// TwinCAT 3 PLC project PLC_Tank
// ProgramVersion: 3.1.4026.27
// libraries:
//   Tc2_ControllerToolbox, * (Beckhoff Automation GmbH)
//   Tc2_ModbusSrv, * (Beckhoff Automation GmbH)
//   Tc2_Standard, * (Beckhoff Automation GmbH)
//   Tc2_System, * (Beckhoff Automation GmbH)
//   Tc3_Module, * (Beckhoff Automation GmbH)
//   VisuDialogs, * (System)
//   VisuSymbols,newest,System
// project tree:
//   DUTs/ TAnalogConversion.TcDUT, TEngine.TcDUT, TEngineCmd.TcDUT, THeaterState.TcDUT, THeaterCmd.TcDUT, THeater.TcDUT, TPhaseHeating.TcDUT, TPhaseCmd.TcDUT, TPhaseDraining.TcDUT, TPhaseFilling.TcDUT, TPhaseMixing.TcDUT, TPhaseState.TcDUT, TValveState.TcDUT, TValveCmd.TcDUT, TEngineState.TcDUT, TTank.TcDUT, TValve.TcDUT
//   / GlobalTextList.TcGTLO, PlcTask.TcTTO, PlcTask500ms.TcTTO, Visualization Manager.TcVMO (not stored)
//   GVLs/ Global.TcGVL
//   POUs/ Draining.TcPOU, Engine_1DO.TcPOU, FB_Tank.TcPOU, Filling.TcPOU, Heater.TcPOU, Heating.TcPOU, Main_Batch.TcPOU, MB_Connector.TcPOU, Mixing.TcPOU, Test.TcPOU, Valve_2DO.TcPOU, MAIN.TcPOU
//   POUs/Misc/ EngToRaw.TcPOU, RawToEng.TcPOU
//   VISUs/ Visualization.TcVIS
// real-time tasks:
//   TASK PlcTask: cycle T#100000us, priority 20, ADS port 350
//   TASK PlcTask500ms: cycle T#500ms, priority 1, ADS port 351

CONFIGURATION PLC_Tank
    RESOURCE PLC ON TwinCAT3
        TASK PlcTask(INTERVAL := T#100000us, PRIORITY := 20);
        TASK PlcTask500ms(INTERVAL := T#500ms, PRIORITY := 1);
        PROGRAM MB_Connector WITH PlcTask : MB_Connector;
        PROGRAM Main_Batch WITH PlcTask : Main_Batch;
        PROGRAM MAIN WITH PlcTask500ms : MAIN;
    END_RESOURCE
END_CONFIGURATION

// ---- DUTs/TAnalogConversion.TcDUT
TYPE TAnalogConversion :
STRUCT
	TransducerLoLevel : UINT;
	TransducerHiLevel : UINT;
	ScaledValLoLevel : REAL;
	ScaledValHiLevel : REAL;
END_STRUCT
END_TYPE

// ---- DUTs/TEngine.TcDUT
TYPE TEngine :
STRUCT
	Cmd : TEngineCmd;
	State : TEngineState;
	Time2Start : TIME := T#5S;
	RisingEdgeTrigger : R_TRIG;
	StartupFailTimer : TON;
END_STRUCT
END_TYPE

// ---- DUTs/TEngineCmd.TcDUT
TYPE TEngineCmd :
STRUCT
		SetRT : DINT;
		AutCtrl : BOOL;
		ManCtrl : BOOL;
		TurnOnMan : BOOL;
		TurnOffMan : BOOL;
		Req2RunAutCtrl : BOOL;
		ResetSUF : BOOL;
END_STRUCT
END_TYPE

// ---- DUTs/THeaterState.TcDUT
TYPE THeaterState :
STRUCT
	EnableOut : BOOL;
	HeatingOut : REAL;
	AutCtrl : BOOL;
	ManCtrl : BOOL;
	MayRun : BOOL;
	MayAutoRun : BOOL;
	Err 	: BOOL;
	StateInt : INT;
	GenErr : BOOL; //signalisation: error occured

	HeatingPower : REAL;
	

END_STRUCT
END_TYPE

// ---- DUTs/THeaterCmd.TcDUT
TYPE THeaterCmd :
STRUCT
	AutCtrl : BOOL;
	ManCtrl : BOOL;
	TurnOnMan : BOOL;
	TurnOffMan : BOOL;
	Req2RunAutCtrl : BOOL;
END_STRUCT
END_TYPE

// ---- DUTs/THeater.TcDUT
TYPE THeater :
STRUCT
	Cmd : THeaterCmd;
	State : THeaterState;
	
	ParamHeatingPowerManual : REAL := 50.0;
	ParamHeatingSetPointAutomat : REAL := 60.0;
	
	PID : FB_CTRL_PID;
	ThresholdTimer : TON;
	
END_STRUCT
END_TYPE

// ---- DUTs/TPhaseHeating.TcDUT
TYPE TPhaseHeating :
STRUCT
	Cmd : TPhaseCmd;
	State : TPhaseState;
	
	ParamReqTemp : REAL;
	
	WaterTemp : REAL;
	
	fTime : INT;
END_STRUCT
END_TYPE

// ---- DUTs/TPhaseCmd.TcDUT
TYPE TPhaseCmd :
STRUCT
	StartAut : BOOL;
	StopAut : BOOL;
	StartMan : BOOL;
	StopMan : BOOL;
	PauseMan : BOOL;
	ResumeMan : BOOL;
	ResetDone : BOOL;
	AutCtrl : BOOL;
	ManCtrl : BOOL;
END_STRUCT
END_TYPE

// ---- DUTs/TPhaseDraining.TcDUT
TYPE TPhaseDraining :
STRUCT
	Cmd : TPhaseCmd;
	State : TPhaseState;
	
	ParamDrainLevel : REAL;
	WaterLevel : REAL;
END_STRUCT
END_TYPE

// ---- DUTs/TPhaseFilling.TcDUT
TYPE TPhaseFilling :
STRUCT
	Cmd : TPhaseCmd;
	State : TPhaseState;
	
	ParamFillLevel : REAL;
	WaterLevel : REAL;
END_STRUCT
END_TYPE

// ---- DUTs/TPhaseMixing.TcDUT
TYPE TPhaseMixing :
STRUCT
	Cmd : TPhaseCmd;
	State : TPhaseState;
	
	ParamTimeSec : INT;
	
	ElapsedTimeSec : INT;
END_STRUCT
END_TYPE

// ---- DUTs/TPhaseState.TcDUT
TYPE TPhaseState :
STRUCT
	Running : BOOL;
	Idle : BOOL;
	Paused : BOOL;
	Done : BOOL;
	AutCtrl : BOOL;
	ManCtrl : BOOL;
	Stateint : INT;
END_STRUCT
END_TYPE

// ---- DUTs/TValveState.TcDUT
TYPE TValveState :
STRUCT
		Open : BOOL;
		Closed : BOOL;
		OpenOut : BOOL;
		CloseOut : BOOL;
		Err : BOOL;
		StartupFail : BOOL;
		AutCtrl : BOOL;
		ManCtrl : BOOL;
		MayRun : BOOL;
		MayAutoRun : BOOL; //device is working in automatic regime
		GenErr : BOOL; //signalisation: error occured
		StColor : INT; //valve state: Open(0), Closed(1), OpenAndErr(2), ClosedAndErr(3) ,NotOpenNotClosedNotErr(4), NotOpenNotClosedAndErr(5), OpenAndClosedAndErr(6), OpenAndClosedNotErr(7)

END_STRUCT
END_TYPE

// ---- DUTs/TValveCmd.TcDUT
TYPE TValveCmd :
STRUCT
		AutCtrl : BOOL;
		ManCtrl : BOOL;
		OpenMan : BOOL;
		StopMan : BOOL;
		CloseMan : BOOL;
		Req2OpenAut : BOOL;
		Req2CloseAut : BOOL;
		ResetSUF : BOOL;
END_STRUCT
END_TYPE

// ---- DUTs/TEngineState.TcDUT
TYPE TEngineState :
STRUCT
		RT : DINT;
		Run : BOOL;
		RunOut : BOOL;
		Err : BOOL;
		StartUpFail : BOOL;
		AutCtrl : BOOL;
		ManCtrl : BOOL;
		MayRun : BOOL;
		MayAutoRun : BOOL;
		GenErr : BOOL;
		StateInt : INT;
		
		StartupFailTime : INT;
END_STRUCT
END_TYPE

// ---- DUTs/TTank.TcDUT
TYPE TTank :
STRUCT
	Mixer : TEngine;
	ValveFilling : TValve;
	ValveDraining : TValve;
	Heater : THeater;
	
	Filling : TPhaseFilling;
	Draining : TPhaseDraining;
	Mixing : TPhaseMixing;
	Heating : TPhaseHeating;
	
	GlobalError : BOOL;

END_STRUCT
END_TYPE

// ---- DUTs/TValve.TcDUT
TYPE TValve :
STRUCT
	Cmd : TValveCmd;
	State : TValveState;
	Time2Open : TIME := T#12S;
	
	OpenFailTimer : TON;
	CloseFailTimer : TON;
	
END_STRUCT
END_TYPE

// ---- GVLs/Global.TcGVL
{attribute 'qualified_only'}
VAR_GLOBAL
	Tank1 : TTank;
	

	secImp : BOOL;
	
	diMixerRun : BOOL;
	diMixerError : BOOL;
	diValveFillOpen : BOOL;
	diValveFillClose : BOOL;
	diValveFillError : BOOL;
	diValveDrainOpen : BOOL;
	diValveDrainClose : BOOL;
	diValveDrainError : BOOL;
	
	aiWaterLevel : WORD;
	aiWaterTemp : WORD;
	
	doMixerStart : BOOL;
	doValveFillOpen : BOOL;
	doValveFillClose : BOOL;
	doValveDrainOpen : BOOL;
	doValveDrainClose : BOOL;
	doHeatingEnable : BOOL;
	
	aoReqPowerOfHeating : WORD;

END_VAR

VAR_GLOBAL CONSTANT
	Running : INT := 0;
	Stop : INT := 1;
	RunningAndError : INT := 2;
	Err : INT := 3;

	PhIdle : INT := 0;
	PhRunning : INT := 1;
	PhPause : INT := 2;
	
    Open : INT := 0;
	Closed : INT := 1;
	OpenAndErr : INT := 2;
	ClosedAndErr : INT := 3;
	NotOpenNotClosedNotErr : INT := 4;
	NotOpenNotClosedAndErr : INT := 5;
	OpenAndClosedAndErr : INT := 6;
	OpenAndClosedNotErr : INT := 7;
END_VAR

// ---- POUs/MB_Connector.TcPOU
PROGRAM MB_Connector
VAR
	
    mb_ipaddr   : STRING(15) := '127.0.0.1';
    mb_port     : UINT := 504;
    mb_unitid   : BYTE := 1;
	
	fbReadRegs		: FB_MBReadInputRegs;
	mb_regs    		: ARRAY [0..4] OF WORD;
	mb_regs_error	: BOOL;
	mb_regs_busy	: BOOL;
	mb_regs_execute : BOOL;
	mb_regs_errid	: UDINT;
	
	fbReadInps	: FB_MBReadInputs;
	mb_inps			: ARRAY [0..4] OF BYTE;
	mb_inps_error	: BOOL;
	mb_inps_busy	: BOOL;
	mb_inps_execute : BOOL;
	mb_inps_errid	: UDINT;
	
	fbWriteRegs		: FB_MBWriteRegs;
	mbw_regs    	: ARRAY [0..4] OF WORD;
	mbw_regs_error	: BOOL;
	mbw_regs_busy	: BOOL;
	mbw_regs_execute: BOOL;
	mbw_regs_errid	: UDINT;
	
	fbWriteCoils	: FB_MBWriteCoils;
	mbw_coils		: ARRAY [0..4] OF BYTE;
	mbw_coils_error	: BOOL;
	mbw_coils_busy	: BOOL;
	mbw_coils_execute: BOOL;
	mbw_coils_errid	: UDINT;
	
END_VAR

fbReadRegs.sIPAddr := mb_ipaddr;
fbReadRegs.nTCPPort := mb_port;
fbReadRegs.nQuantity := 4;
fbReadRegs.nMBAddr := 0;
fbReadRegs.cbLength := SIZEOF(mb_regs);
fbReadRegs.pDestAddr := ADR(mb_regs);
fbReadRegs.nUnitID := mb_unitid;
fbReadRegs.tTimeout := T#5S;
IF (mb_regs_busy = FALSE) THEN
	mb_regs_execute := TRUE;
ELSE
	mb_regs_execute := FALSE;
END_IF
fbReadRegs(bExecute := mb_regs_execute, 
		   bBusy => mb_regs_busy, bError => mb_regs_error, 
		   nErrId => mb_regs_errid);



fbReadInps.sIPAddr := mb_ipaddr;
fbReadInps.nTCPPort := mb_port;
fbReadInps.nQuantity := 32;
fbReadInps.nMBAddr := 0;
fbReadInps.cbLength := SIZEOF(mb_inps);
fbReadInps.pDestAddr := ADR(mb_inps);
fbReadInps.nUnitID := mb_unitid;
fbReadInps.tTimeout := T#5S;
IF (mb_inps_busy = FALSE) THEN
	mb_inps_execute := TRUE;
ELSE
	mb_inps_execute := FALSE;
END_IF
fbReadInps(bExecute := mb_inps_execute, 
	bBusy => mb_inps_busy, bError => mb_inps_error, nErrId => mb_inps_errid);

Global.diValveFillOpen := mb_inps[0].0;
Global.diValveFillClose := mb_inps[0].1;
Global.diValveFillError := mb_inps[0].2;
Global.diValveDrainOpen := mb_inps[0].3;
Global.diValveDrainClose := mb_inps[0].4;
Global.diValveDrainError := mb_inps[0].5;
Global.diMixerRun := mb_inps[0].6;
Global.diMixerError := mb_inps[0].7;

Global.aiWaterLevel := mb_regs[0];
Global.aiWaterTemp := mb_regs[2];







fbWriteRegs.sIPAddr := mb_ipaddr;
fbWriteRegs.nTCPPort := mb_port;
fbWriteRegs.nQuantity := 4;
fbWriteRegs.nMBAddr := 0;
fbWriteRegs.cbLength := SIZEOF(mbw_regs);
fbWriteRegs.pSrcAddr := ADR(mbw_regs);
fbWriteRegs.nUnitID := mb_unitid;
fbWriteRegs.tTimeout := T#5S;
IF (mbw_regs_busy = FALSE) THEN
	mbw_regs_execute := TRUE;
ELSE
	mbw_regs_execute := FALSE;
END_IF
fbWriteRegs(bExecute := mbw_regs_execute, 
		   bBusy => mbw_regs_busy, bError => mbw_regs_error, 
		   nErrId => mbw_regs_errid);



fbWriteCoils.sIPAddr := mb_ipaddr;
fbWriteCoils.nTCPPort := mb_port;
fbWriteCoils.nQuantity := 32;
fbWriteCoils.nMBAddr := 0;
fbWriteCoils.cbLength := SIZEOF(mbw_coils);
fbWriteCoils.pSrcAddr := ADR(mbw_coils);
fbWriteCoils.nUnitID := mb_unitid;
fbWriteCoils.tTimeout := T#5S;
IF (mbw_coils_busy = FALSE) THEN
	mbw_coils_execute := TRUE;
ELSE
	mbw_coils_execute := FALSE;
END_IF
fbWriteCoils(bExecute := mbw_coils_execute, 
	bBusy => mbw_coils_busy, bError => mbw_coils_error, nErrId => mbw_coils_errid);

mbw_coils[0].0 := Global.doValveFillOpen;
mbw_coils[0].1 := Global.doValveFillClose;
mbw_coils[0].2 := Global.doValveDrainOpen;
mbw_coils[0].3 := Global.doValveDrainClose;
mbw_coils[0].4 := Global.doMixerStart;
mbw_coils[0].5 := Global.doHeatingEnable;

mbw_regs[0] := Global.aoReqPowerOfHeating;

END_PROGRAM

// ---- POUs/Main_Batch.TcPOU
PROGRAM Main_Batch
VAR
	FB_Tank_1 : FB_Tank;
END_VAR

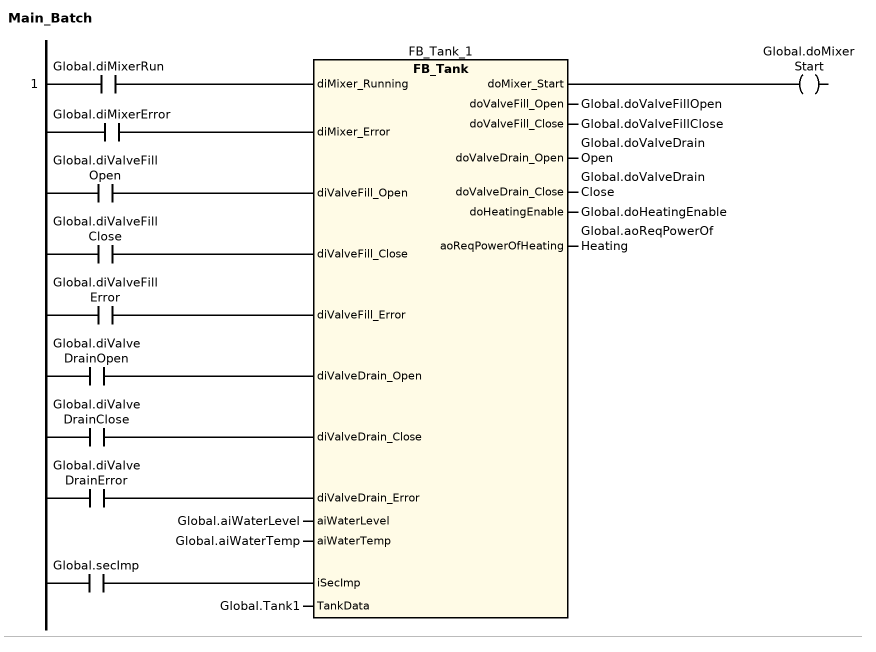
// NETWORK 1
FB_Tank_1(
    diMixer_Running := Global.diMixerRun,
    diMixer_Error := Global.diMixerError,
    diValveFill_Open := Global.diValveFillOpen,
    diValveFill_Close := Global.diValveFillClose,
    diValveFill_Error := Global.diValveFillError,
    diValveDrain_Open := Global.diValveDrainOpen,
    diValveDrain_Close := Global.diValveDrainClose,
    diValveDrain_Error := Global.diValveDrainError,
    aiWaterLevel := Global.aiWaterLevel,
    aiWaterTemp := Global.aiWaterTemp,
    iSecImp := Global.secImp,
    TankData := Global.Tank1,
    doValveFill_Open => Global.doValveFillOpen,
    doValveFill_Close => Global.doValveFillClose,
    doValveDrain_Open => Global.doValveDrainOpen,
    doValveDrain_Close => Global.doValveDrainClose,
    doHeatingEnable => Global.doHeatingEnable,
    aoReqPowerOfHeating => Global.aoReqPowerOfHeating); // FB_Tank
Global.doMixerStart := FB_Tank_1.doMixer_Start;

END_PROGRAM

// ---- POUs/FB_Tank.TcPOU
FUNCTION_BLOCK FB_Tank
VAR_INPUT
	diMixer_Running : BOOL;
	diMixer_Error : BOOL;
	diValveFill_Open : BOOL;
	diValveFill_Close : BOOL;
	diValveFill_Error : BOOL;
	diValveDrain_Open : BOOL;
	diValveDrain_Close : BOOL;
	diValveDrain_Error : BOOL;
	aiWaterLevel : WORD;
	aiWaterTemp : WORD;
	iSecImp : BOOL; //Požaduje se vstup s periodou 1 sekunda a libovolnou střídou
END_VAR

VAR_OUTPUT
	doMixer_Start : BOOL;
	doValveFill_Open : BOOL;
	doValveFill_Close : BOOL;
	doValveDrain_Open : BOOL;
	doValveDrain_Close : BOOL;
	doHeatingEnable : BOOL;
	aoReqPowerOfHeating : WORD;
END_VAR

VAR_IN_OUT
	TankData : TTank;
END_VAR

VAR
	//Konfigurace přepočtu rozsahu převodníků
	WaterTemp : TAnalogConversion := (TransducerLoLevel := 0, TransducerHiLevel := 27648, ScaledValLoLevel := 0, ScaledValHiLevel := 100);
	WaterLevel : TAnalogConversion := (TransducerLoLevel := 0, TransducerHiLevel := 27648, ScaledValLoLevel := 0, ScaledValHiLevel := 2);
	ReqOutputPower : TAnalogConversion := (ScaledValLoLevel := 0, ScaledValHiLevel := 100, TransducerLoLevel := 0, TransducerHiLevel := 27648);

	//Instance zanořených funkčních bloků
	ValveDrainCm : Valve_2DO;
	ValveFillCm : Valve_2DO;
	MixerCm : Engine_1DO;
	HeaterCm : Heater;
	FillingPhase : Filling;
	MixingPhase : Mixing;
	DrainingPhase : Draining;
	HeatingPhase : Heating;
	TON1: TON;
	RawToEng_1: RawToEng;
	RawToEng_2: RawToEng;
	EngToRaw_1: EngToRaw;
END_VAR

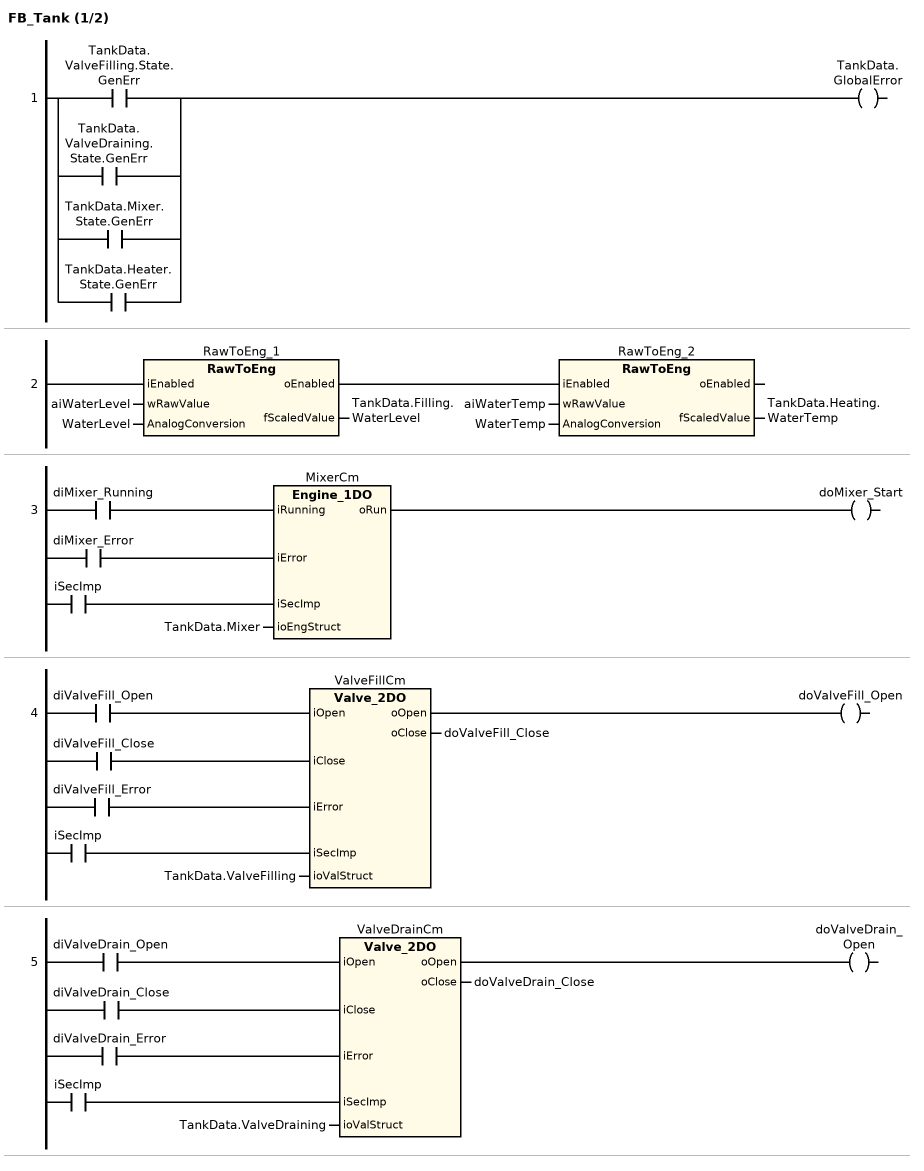
// NETWORK 1
TankData.GlobalError := TankData.ValveFilling.State.GenErr OR TankData.ValveDraining.State.GenErr OR TankData.Mixer.State.GenErr OR TankData.Heater.State.GenErr;

// NETWORK 2
RawToEng_1(
    iEnabled := TRUE,
    wRawValue := aiWaterLevel,
    AnalogConversion := WaterLevel,
    fScaledValue => TankData.Filling.WaterLevel); // RawToEng
RawToEng_2(
    iEnabled := RawToEng_1.oEnabled,
    wRawValue := aiWaterTemp,
    AnalogConversion := WaterTemp,
    fScaledValue => TankData.Heating.WaterTemp); // RawToEng

// NETWORK 3
MixerCm(
    iRunning := diMixer_Running,
    iError := diMixer_Error,
    iSecImp := iSecImp,
    ioEngStruct := TankData.Mixer); // Engine_1DO
doMixer_Start := MixerCm.oRun;

// NETWORK 4
ValveFillCm(
    iOpen := diValveFill_Open,
    iClose := diValveFill_Close,
    iError := diValveFill_Error,
    iSecImp := iSecImp,
    ioValStruct := TankData.ValveFilling,
    oClose => doValveFill_Close); // Valve_2DO
doValveFill_Open := ValveFillCm.oOpen;

// NETWORK 5
ValveDrainCm(
    iOpen := diValveDrain_Open,
    iClose := diValveDrain_Close,
    iError := diValveDrain_Error,
    iSecImp := iSecImp,
    ioValStruct := TankData.ValveDraining,
    oClose => doValveDrain_Close); // Valve_2DO
doValveDrain_Open := ValveDrainCm.oOpen;

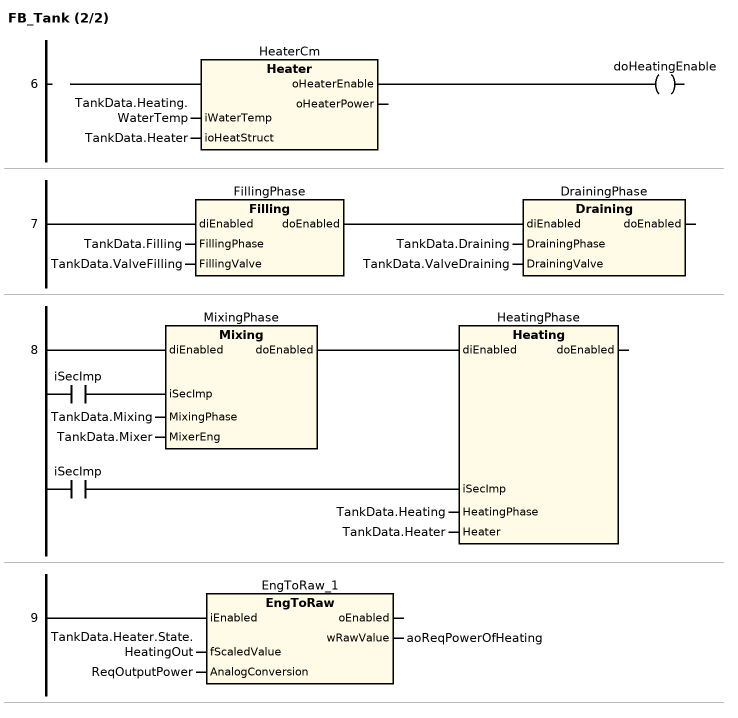
// NETWORK 6
HeaterCm(iWaterTemp := TankData.Heating.WaterTemp, ioHeatStruct := TankData.Heater); // Heater
doHeatingEnable := HeaterCm.oHeaterEnable;

// NETWORK 7
FillingPhase(diEnabled := TRUE, FillingPhase := TankData.Filling, FillingValve := TankData.ValveFilling); // Filling
DrainingPhase(
    diEnabled := FillingPhase.doEnabled,
    DrainingPhase := TankData.Draining,
    DrainingValve := TankData.ValveDraining); // Draining

// NETWORK 8
MixingPhase(
    diEnabled := TRUE,
    iSecImp := iSecImp,
    MixingPhase := TankData.Mixing,
    MixerEng := TankData.Mixer); // Mixing
HeatingPhase(
    diEnabled := MixingPhase.doEnabled,
    iSecImp := iSecImp,
    HeatingPhase := TankData.Heating,
    Heater := TankData.Heater); // Heating

// NETWORK 9
EngToRaw_1(
    iEnabled := TRUE,
    fScaledValue := TankData.Heater.State.HeatingOut,
    AnalogConversion := ReqOutputPower,
    wRawValue => aoReqPowerOfHeating); // EngToRaw

END_FUNCTION_BLOCK

// ---- POUs/Valve_2DO.TcPOU
FUNCTION_BLOCK Valve_2DO
VAR_INPUT
	iOpen : BOOL;
	iClose : BOOL;
	iError : BOOL;
	iSecImp : BOOL;
END_VAR
VAR_OUTPUT
	oOpen : BOOL;
	oClose : BOOL;
END_VAR

VAR_IN_OUT
	ioValStruct	 : TValve;
END_VAR

VAR
	tempOpenStartupFail : BOOL;
	tempCloseStartupFail: BOOL;
END_VAR

{region "OpenState"}
    // set real state of valve input into valve structure - input of valve can be taken from limit sensor...
    ioValStruct.State.Open := iOpen;
    ioValStruct.State.Closed := iClose;
{endregion}

	 
{region "Manual/Automat"}
	// switching state of engine - automatic or manual control (default state is manual)
	IF ioValStruct.Cmd.ManCtrl THEN
		ioValStruct.State.ManCtrl := TRUE;
		ioValStruct.State.AutCtrl := FALSE;
	ELSIF ioValStruct.Cmd.AutCtrl THEN
		ioValStruct.State.ManCtrl := FALSE;
		ioValStruct.State.AutCtrl := TRUE;
	END_IF;

	IF (NOT ioValStruct.State.ManCtrl) AND (NOT ioValStruct.State.AutCtrl) THEN
		ioValStruct.State.ManCtrl := TRUE;
		ioValStruct.State.AutCtrl := FALSE;
	END_IF;

	ioValStruct.Cmd.ManCtrl := FALSE;
	ioValStruct.Cmd.AutCtrl := FALSE;
{endregion}
	 
{region "MayRun / MayAutoRun"}
    // setting auxilary signals (may run, may auto run) - MR AND NOT MAR - engine may be started in manual mode, MAR - engine may be started in automatic mode
    ioValStruct.State.MayRun := (ioValStruct.State.ManCtrl AND NOT(ioValStruct.State.GenErr));
	ioValStruct.State.MayAutoRun := (ioValStruct.State.AutCtrl AND NOT(ioValStruct.State.GenErr));
{endregion}
	 
{region "ManCtrl"}
	// processing manual actions - if command is processed, it is sets to FALSE even if can't be processed
    // Valve commands are open, close and stop - valve can be stopped intermediate position
	 IF ioValStruct.State.ManCtrl AND ioValStruct.State.MayRun THEN
        IF ioValStruct.Cmd.OpenMan THEN
            ioValStruct.State.CloseOut := FALSE;
            ioValStruct.State.OpenOut := TRUE;
        END_IF;
        
        IF ioValStruct.Cmd.CloseMan THEN
            ioValStruct.State.OpenOut := FALSE;
            ioValStruct.State.CloseOut := TRUE;
        END_IF;
        
        IF ioValStruct.Cmd.StopMan THEN
            ioValStruct.State.OpenOut := FALSE;
            ioValStruct.State.CloseOut := FALSE;
        END_IF;
    END_IF;
    
    ioValStruct.Cmd.OpenMan := FALSE;
    ioValStruct.Cmd.CloseMan := FALSE;
    ioValStruct.Cmd.StopMan := FALSE;
{endregion}
	 
{region "AutCtrl"}
	 //if request to run in automatic mode -> set outputs to right states if MAR
    //AutoRequest shouldn't be reseted to false state
    //if request to open and request to close are setted to 1 simultaneously - outputs should be 0.
    IF ioValStruct.State.AutCtrl AND ioValStruct.State.MayAutoRun THEN
        IF ioValStruct.Cmd.Req2CloseAut AND (NOT ioValStruct.Cmd.Req2OpenAut) THEN
            ioValStruct.State.OpenOut := FALSE;
            ioValStruct.State.CloseOut := TRUE;
        ELSIF (NOT ioValStruct.Cmd.Req2CloseAut) AND ioValStruct.Cmd.Req2OpenAut THEN
            ioValStruct.State.CloseOut := FALSE;
            ioValStruct.State.OpenOut := TRUE;
        ELSE
            ioValStruct.State.CloseOut := FALSE;
            ioValStruct.State.OpenOut := FALSE;
        END_IF;
        
    END_IF;
{endregion}
	 
{region "Error states"}
 // definition of error states 
    // error - input from digital input of plc - fyzical state of valve
    // calculating start up fail - if output is sets to open or close, it's expected feedback from limit sensor in defined time, if feedback doesn't show in this time, it should be start up fail error
    // merge of these two error is general error
    // error is both inputs (open and closed) true state
    ioValStruct.OpenFailTimer(IN := (ioValStruct.State.OpenOut AND (NOT ioValStruct.State.CloseOut) AND (NOT ioValStruct.State.Open)), PT := ioValStruct.Time2Open);
	tempOpenStartupFail := ioValStruct.OpenFailTimer.Q;

    ioValStruct.CloseFailTimer(IN := ((NOT ioValStruct.State.OpenOut) AND ioValStruct.State.CloseOut AND (NOT ioValStruct.State.Closed)), PT := ioValStruct.Time2Open);
	tempCloseStartupFail := ioValStruct.CloseFailTimer.Q;
    
   
    IF tempOpenStartupFail OR tempCloseStartupFail THEN
        ioValStruct.State.StartupFail := TRUE;
    END_IF;
    
    ioValStruct.State.Err := iError OR (ioValStruct.State.Open AND ioValStruct.State.Closed);
    
    // start up fail can be reseted by operator, command resetSUF, resets SUF and engine should be started again
    IF ioValStruct.Cmd.ResetSUF THEN
        ioValStruct.State.StartupFail := FALSE;
        ioValStruct.Cmd.ResetSUF := FALSE;
    END_IF;

    ioValStruct.State.GenErr := ioValStruct.State.StartupFail OR ioValStruct.State.Err;
    
    // if error state exists outputs should be in stop state
    IF ioValStruct.State.GenErr THEN
        ioValStruct.State.OpenOut := FALSE;
        ioValStruct.State.CloseOut := FALSE;
    END_IF;
{endregion}
	 	 
oOpen := ioValStruct.State.OpenOut;
oClose := ioValStruct.State.CloseOut;

{region "StatusInt"}
    //write combination of states into int value for visualization (valve - combination of open, close state and error)
    IF ioValStruct.State.Open AND NOT ioValStruct.State.Closed AND NOT ioValStruct.State.GenErr THEN
        ioValStruct.State.StColor := Global.Open;
    ELSIF NOT ioValStruct.State.Open AND ioValStruct.State.Closed AND NOT ioValStruct.State.GenErr THEN
        ioValStruct.State.StColor := Global.Closed;
    ELSIF ioValStruct.State.Open AND NOT ioValStruct.State.Closed AND ioValStruct.State.GenErr THEN
        ioValStruct.State.StColor := Global.OpenAndErr;
    ELSIF NOT ioValStruct.State.Open AND ioValStruct.State.Closed AND ioValStruct.State.GenErr THEN
        ioValStruct.State.StColor := Global.ClosedAndErr;
    ELSIF NOT ioValStruct.State.Open AND NOT ioValStruct.State.Closed AND NOT ioValStruct.State.GenErr THEN
        ioValStruct.State.StColor := Global.NotOpenNotClosedNotErr;
    ELSIF NOT ioValStruct.State.Open AND NOT ioValStruct.State.Closed AND ioValStruct.State.GenErr THEN
        ioValStruct.State.StColor := Global.NotOpenNotClosedAndErr;
    ELSIF ioValStruct.State.Open AND ioValStruct.State.Closed AND ioValStruct.State.GenErr THEN
        ioValStruct.State.StColor := Global.OpenAndClosedAndErr;
    ELSIF ioValStruct.State.Open AND ioValStruct.State.Closed AND NOT ioValStruct.State.GenErr THEN
        ioValStruct.State.StColor := Global.OpenAndClosedNotErr;
    END_IF;
{endregion}

END_FUNCTION_BLOCK

// ---- POUs/Engine_1DO.TcPOU
FUNCTION_BLOCK Engine_1DO
VAR_INPUT
	iRunning : BOOL;
	iError : BOOL;
	iSecImp : BOOL;
END_VAR
VAR_OUTPUT
	oRun : BOOL;
END_VAR
VAR_IN_OUT
	ioEngStruct : TEngine;
END_VAR
VAR
	secImpEdge: BOOL;
	tempStartupFail: BOOL;
END_VAR

{region "RunState"}
    // set real state of engine run into engine structure
    ioEngStruct.State.Run := iRunning;
{endregion}

{region "Running time"} 
    // counting running time of engine - (motoseconds in real situation it should be moto hours)
    // detection rising edge of input secimp - should be conected 1Hz internal clock from PLC
	ioEngStruct.RisingEdgeTrigger(CLK := iSecImp, Q => secImpEdge);
	IF ioEngStruct.State.Run AND secImpEdge THEN
		ioEngStruct.State.RT := ioEngStruct.State.RT + 1;
	END_IF;

	IF ioEngStruct.Cmd.SetRT >= 0 THEN
		ioEngStruct.State.RT := ioEngStruct.Cmd.SetRT;
		ioEngStruct.Cmd.SetRT := -1;
	END_IF;
{endregion}
	 
 
{region "Manual/Automat"}
	// switching state of engine - automatic or manual control (default state is manual)
	IF ioEngStruct.Cmd.ManCtrl THEN
		ioEngStruct.State.ManCtrl := TRUE;
		ioEngStruct.State.AutCtrl := FALSE;
	ELSIF ioEngStruct.Cmd.AutCtrl THEN
		ioEngStruct.State.ManCtrl := FALSE;
		ioEngStruct.State.AutCtrl := TRUE;
	END_IF;

	IF (NOT ioEngStruct.State.ManCtrl) AND (NOT ioEngStruct.State.AutCtrl) THEN
		ioEngStruct.State.ManCtrl := TRUE;
		ioEngStruct.State.AutCtrl := FALSE;
	END_IF;

	ioEngStruct.Cmd.ManCtrl := FALSE;
	ioEngStruct.Cmd.AutCtrl := FALSE;
{endregion}
	 
{region "MayRun / MayAutoRun"}
	// setting auxilary signals (may run, may auto run) - MR AND NOT MAR - eng should be started in manual mode,
    // MAR - should be started in automatic mode
    ioEngStruct.State.MayRun := (ioEngStruct.State.ManCtrl AND NOT(ioEngStruct.State.GenErr));
	ioEngStruct.State.MayAutoRun := (ioEngStruct.State.AutCtrl AND NOT(ioEngStruct.State.GenErr));
		 
			  
{endregion}
	 
{region "ManCtrl"}
	// processing manual actions - if command is processed, it is set to FALSE even if can't be processed
    // Engine commands are turn off (stop) and turn on (start)
	IF ioEngStruct.State.ManCtrl AND ioEngStruct.State.MayRun THEN
		IF ioEngStruct.Cmd.TurnOnMan THEN
			ioEngStruct.State.RunOut := TRUE;
		END_IF;

		IF ioEngStruct.Cmd.TurnOffMan THEN
			ioEngStruct.State.RunOut := FALSE;
		END_IF;
	END_IF;

	ioEngStruct.Cmd.TurnOnMan := FALSE;
	ioEngStruct.Cmd.TurnOffMan := FALSE;
{endregion}
	 
{region "AutCtrl"}
	//if request to run in automatic mode set outputs to right states if MAR
    //AutoRequest shouldn't be reseted to false state
    IF ioEngStruct.State.AutCtrl AND ioEngStruct.State.MayAutoRun THEN
		ioEngStruct.State.RunOut := ioEngStruct.Cmd.Req2RunAutCtrl;
	END_IF;
{endregion}
	 
{region "Error states"}
	// definition of error states 
	// error - input from digital input of plc - fyzical state of engine 
	// calculating start up fail - if output is sets to start engine, it's expected feedback from running signal in defined time, if feedback doesn't show in this time, it should be start up fail error
	// merge of these two error is general error
	ioEngStruct.StartupFailTimer(IN := (ioEngStruct.State.RunOut AND (NOT ioEngStruct.State.Run)), PT := ioEngStruct.Time2Start);
	tempStartupFail := ioEngStruct.StartupFailTimer.Q;

	IF tempStartupFail THEN
		ioEngStruct.State.StartUpFail := TRUE;
	END_IF;

	ioEngStruct.State.Err := iError;

	IF ioEngStruct.Cmd.ResetSUF THEN
		ioEngStruct.State.StartUpFail := FALSE;
		ioEngStruct.Cmd.ResetSUF := FALSE;
	END_IF;

	ioEngStruct.State.GenErr := ioEngStruct.State.StartUpFail OR ioEngStruct.State.Err;

	IF ioEngStruct.State.GenErr THEN
		ioEngStruct.State.RunOut := FALSE;
	END_IF;
{endregion}
	 
oRun := ioEngStruct.State.RunOut;

{region "StatusInt"}
 IF NOT ioEngStruct.State.GenErr THEN
        IF ioEngStruct.State.Run THEN
            ioEngStruct.State.StateInt := Global.Running;
        ELSE
            ioEngStruct.State.StateInt := Global.Stop;
        END_IF;
    ELSE
        IF ioEngStruct.State.Run THEN
            ioEngStruct.State.StateInt := Global.RunningAndError;
        ELSE
            ioEngStruct.State.StateInt := Global.Err;
        END_IF;
    END_IF; 
{endregion}

END_FUNCTION_BLOCK

// ---- POUs/Heater.TcPOU
FUNCTION_BLOCK Heater
VAR_INPUT
	iWaterTemp : REAL;
END_VAR
VAR_OUTPUT
	oHeaterEnable : BOOL;
	oHeaterPower : REAL;
END_VAR
VAR_IN_OUT
	ioHeatStruct : THeater;
END_VAR
VAR
	pidParameters : ST_CTRL_PID_PARAMS;
END_VAR

pidParameters.fKp := 10; //P
pidParameters.tTn := T#2S; //I
pidParameters.tTv := T#0.5S; //D
pidParameters.tCtrlCycleTime := T#200MS;
pidParameters.tTaskCycleTime := T#100MS;
pidParameters.fOutMaxLimit := 100;
pidParameters.fOutMinLimit := 0;
pidParameters.bDInTheFeedbackPath := FALSE;
pidParameters.bPInTheFeedbackPath := FALSE;
pidParameters.bARWOnIPartOnly := FALSE;
pidParameters.tTd := T#100MS; 

ioHeatStruct.PID(
	fSetpointValue := ioHeatStruct.ParamHeatingSetPointAutomat, 
	fActualValue := iWaterTemp, 
	fManSyncValue := ioHeatStruct.ParamHeatingPowerManual,
	bSync := ioHeatStruct.State.ManCtrl,
	eMode := E_CTRL_MODE.eCTRL_MODE_ACTIVE, // automatic mode of PID component
	stParams := pidParameters);

ioHeatStruct.State.HeatingOut := ioHeatStruct.PID.fOut;

	 
{region "Manual/Automat"}
// switching state of engine - automatic or manual control (default state is manual)
IF ioHeatStruct.Cmd.ManCtrl THEN
	ioHeatStruct.State.ManCtrl := TRUE;
	ioHeatStruct.State.AutCtrl := FALSE;
ELSIF ioHeatStruct.Cmd.AutCtrl THEN
	ioHeatStruct.State.ManCtrl := FALSE;
	ioHeatStruct.State.AutCtrl := TRUE;
END_IF;

IF (NOT ioHeatStruct.State.ManCtrl) AND (NOT ioHeatStruct.State.AutCtrl) THEN
	ioHeatStruct.State.ManCtrl := TRUE;
	ioHeatStruct.State.AutCtrl := FALSE;
END_IF;

ioHeatStruct.Cmd.ManCtrl := FALSE;
ioHeatStruct.Cmd.AutCtrl := FALSE;

ioHeatStruct.State.MayRun := (ioHeatStruct.State.ManCtrl AND NOT(ioHeatStruct.State.GenErr));
ioHeatStruct.State.MayAutoRun := (ioHeatStruct.State.AutCtrl AND NOT(ioHeatStruct.State.GenErr));
{endregion}
	 
 
{region "ManCtrl"}
// processing manual actions - if command is processed, it is set to FALSE even if can't be processed
// Engine commands are turn off (stop) and turn on (start)
IF ioHeatStruct.State.ManCtrl AND ioHeatStruct.State.MayRun THEN
	IF ioHeatStruct.Cmd.TurnOnMan THEN
		ioHeatStruct.State.EnableOut := TRUE;
	END_IF;

	IF ioHeatStruct.Cmd.TurnOffMan THEN
		ioHeatStruct.State.EnableOut := FALSE;
	END_IF;

	IF ioHeatStruct.State.EnableOut THEN
		ioHeatStruct.State.HeatingOut := LIMIT(0.0, ioHeatStruct.ParamHeatingPowerManual, 100.0);
	ELSE
		ioHeatStruct.State.HeatingOut := 0.0;
	END_IF;
END_IF;

ioHeatStruct.Cmd.TurnOnMan := FALSE;
ioHeatStruct.Cmd.TurnOffMan := FALSE;
{endregion}
 
{region "AutCtrl"}
//if request to run in automatic mode set outputs to right states if MAR
//AutoRequest shouldn't be reseted to false state
IF ioHeatStruct.State.AutCtrl AND ioHeatStruct.State.MayAutoRun THEN
	ioHeatStruct.State.EnableOut := ioHeatStruct.Cmd.Req2RunAutCtrl;

	IF ioHeatStruct.State.EnableOut THEN
		ioHeatStruct.State.HeatingOut := ioHeatStruct.PID.fOut;
	ELSE
		ioHeatStruct.State.HeatingOut := 0.0;
	END_IF;
END_IF;
{endregion}
 
{region "Error states"}
// if water temperature is too high, stop heating and generate error
ioHeatStruct.ThresholdTimer(IN := (iWaterTemp > 95.0), PT := T#2S);
ioHeatStruct.State.Err := ioHeatStruct.ThresholdTimer.Q OR (iWaterTemp >= 98.0);
ioHeatStruct.State.GenErr := ioHeatStruct.State.Err;

IF ioHeatStruct.State.GenErr THEN
	ioHeatStruct.State.EnableOut := FALSE;
	ioHeatStruct.State.HeatingOut := 0.0;
END_IF;

IF NOT ioHeatStruct.State.EnableOut THEN
	ioHeatStruct.State.HeatingOut := 0.0;
END_IF;

ioHeatStruct.State.HeatingPower := ioHeatStruct.State.HeatingOut;

IF NOT ioHeatStruct.State.GenErr THEN
	IF ioHeatStruct.State.EnableOut THEN
		ioHeatStruct.State.StateInt := Global.Running;
	ELSE
		ioHeatStruct.State.StateInt := Global.Stop;
	END_IF;
ELSE
	IF ioHeatStruct.State.EnableOut THEN
		ioHeatStruct.State.StateInt := Global.RunningAndError;
	ELSE
		ioHeatStruct.State.StateInt := Global.Err;
	END_IF;
END_IF;
{endregion}
	 
 
oHeaterPower := ioHeatStruct.State.HeatingOut;
oHeaterEnable := ioHeatStruct.State.EnableOut;

END_FUNCTION_BLOCK

// ---- POUs/Filling.TcPOU
FUNCTION_BLOCK Filling
VAR_INPUT
	diEnabled : BOOL;
END_VAR
VAR_OUTPUT
	doEnabled : BOOL;
END_VAR
VAR_IN_OUT
	FillingPhase : TPhaseFilling;
	FillingValve : TValve;
END_VAR
VAR
END_VAR

{region "REGION Aut/Man"}
    // switching state of engine - automatic or manual control (default state is manual)
    IF FillingPhase.Cmd.ManCtrl THEN
        FillingPhase.State.ManCtrl := TRUE;
        FillingPhase.State.AutCtrl := FALSE;
    ELSIF FillingPhase.Cmd.AutCtrl THEN
        FillingPhase.State.ManCtrl := FALSE;
        FillingPhase.State.AutCtrl := TRUE;
    END_IF;

    IF (NOT FillingPhase.State.ManCtrl) AND (NOT FillingPhase.State.AutCtrl) THEN
        FillingPhase.State.ManCtrl := TRUE;
        FillingPhase.State.AutCtrl := FALSE;
    END_IF;

    FillingPhase.Cmd.ManCtrl := FALSE;
    FillingPhase.Cmd.AutCtrl := FALSE;
{endregion}

{region "ManCtrl"}
    // processing manual actions - if command is processed, it is sets to FALSE even if can't be processed
    // Phase commands are start, stop, pause and resume 
    // Start - open filling valve 
    // Stop - close filling valve
    // Pause - close filling valve
    // Resume - open filling valve
    // real states of phase are writed into states in phase structure
    IF FillingPhase.State.ManCtrl THEN
        IF FillingPhase.Cmd.StartMan THEN
            FillingPhase.State.Done := FALSE;
            IF FillingPhase.State.Idle THEN
                FillingPhase.State.Idle    := FALSE;
                FillingPhase.State.Paused  := FALSE;
                FillingPhase.State.Running := TRUE;
            END_IF;
        END_IF;

        IF FillingPhase.Cmd.PauseMan THEN
            FillingPhase.State.Done := FALSE;
            IF FillingPhase.State.Running THEN
                FillingPhase.State.Running := FALSE;
                FillingPhase.State.Idle    := FALSE;
                FillingPhase.State.Paused  := TRUE;
            END_IF;
        END_IF;

        IF FillingPhase.Cmd.ResumeMan THEN
            FillingPhase.State.Done := FALSE;
            IF FillingPhase.State.Paused THEN
                FillingPhase.State.Paused  := FALSE;
                FillingPhase.State.Idle    := FALSE;
                FillingPhase.State.Running := TRUE;
            END_IF;
        END_IF;

        IF FillingPhase.Cmd.StopMan THEN
            FillingPhase.State.Done    := FALSE;
            FillingPhase.State.Running := FALSE;
            FillingPhase.State.Paused  := FALSE;
            FillingPhase.State.Idle    := TRUE;
        END_IF;
    END_IF;

    FillingPhase.Cmd.StartMan  := FALSE;
    FillingPhase.Cmd.StopMan   := FALSE;
    FillingPhase.Cmd.PauseMan  := FALSE;
    FillingPhase.Cmd.ResumeMan := FALSE;
{endregion}

{region "AutCtrl"}
    // if request to run in automatic mode and phase can be run in automatic mode switch phase to running
    IF FillingPhase.State.AutCtrl THEN
        IF FillingPhase.Cmd.StartAut THEN
            FillingPhase.State.Done := FALSE;
            IF FillingPhase.State.Idle THEN
                FillingPhase.State.Idle    := FALSE;
                FillingPhase.State.Paused  := FALSE;
                FillingPhase.State.Running := TRUE;
            END_IF;
        END_IF;

        IF FillingPhase.Cmd.StopAut THEN
            FillingPhase.State.Done    := FALSE;
            FillingPhase.State.Running := FALSE;
            FillingPhase.State.Paused  := FALSE;
            FillingPhase.State.Idle    := TRUE;
        END_IF;
    END_IF;

    FillingPhase.Cmd.StartAut := FALSE;
    FillingPhase.Cmd.StopAut  := FALSE;
{endregion}

{region "Done"}
    //every phase should have finish condition - filling phase - if water level is above requested level
    //after that done state should be setted to 1
    IF FillingPhase.State.Running THEN
        IF FillingPhase.WaterLevel >= FillingPhase.ParamFillLevel THEN
            FillingPhase.State.Running := FALSE;
            FillingPhase.State.Paused  := FALSE;
            FillingPhase.State.Idle    := TRUE;
            FillingPhase.State.Done    := TRUE;
        END_IF;
    END_IF;

    IF FillingPhase.Cmd.ResetDone THEN
        FillingPhase.State.Done    := FALSE;
        FillingPhase.Cmd.ResetDone := FALSE;
    END_IF;
{endregion}

{region "States"} 
    //Command valve in cases of states
    IF FillingPhase.State.Running THEN
        FillingValve.Cmd.Req2OpenAut  := TRUE;
        FillingValve.Cmd.Req2CloseAut := FALSE;
    ELSE
        FillingValve.Cmd.Req2OpenAut  := FALSE;
        FillingValve.Cmd.Req2CloseAut := TRUE;
    END_IF;
{endregion}


// delault state of phase - if not any state sets state to idle
IF NOT FillingPhase.State.Idle AND NOT FillingPhase.State.Paused AND NOT FillingPhase.State.Running THEN
    FillingPhase.State.Idle := 1;
END_IF;

// write binary states into int value for visualization
IF FillingPhase.State.Idle THEN
    FillingPhase.State.Stateint := Global.PhIdle;
ELSIF FillingPhase.State.Running THEN
    FillingPhase.State.Stateint := Global.PhRunning;
ELSE
    FillingPhase.State.Stateint := Global.PhPause;
END_IF;

// Ponechte pro moznost retezeni volani bloku v LAD
doEnabled := diEnabled;

END_FUNCTION_BLOCK

// ---- POUs/Mixing.TcPOU
FUNCTION_BLOCK Mixing
VAR_INPUT
	diEnabled : BOOL;
	iSecImp : BOOL;
END_VAR
VAR_OUTPUT
	doEnabled : BOOL;
END_VAR
VAR_IN_OUT
	MixingPhase : TPhaseMixing;
	MixerEng : TEngine;
END_VAR
VAR
	secImpTrig : R_TRIG;
END_VAR

{region "Aut/Man"}
    // switching state of engine - automatic or manual control (default state is manual)
    IF MixingPhase.Cmd.ManCtrl THEN
        MixingPhase.State.ManCtrl := TRUE;
        MixingPhase.State.AutCtrl := FALSE;
    ELSIF MixingPhase.Cmd.AutCtrl THEN
        MixingPhase.State.ManCtrl := FALSE;
        MixingPhase.State.AutCtrl := TRUE;
    END_IF;

    IF (NOT MixingPhase.State.ManCtrl) AND (NOT MixingPhase.State.AutCtrl) THEN
        MixingPhase.State.ManCtrl := TRUE;
        MixingPhase.State.AutCtrl := FALSE;
    END_IF;

    MixingPhase.Cmd.ManCtrl := FALSE;
    MixingPhase.Cmd.AutCtrl := FALSE;
{endregion}

{region "ManCtrl"}
    // processing manual actions - if command is processed, it is sets to FALSE even if can't be processed
    // Phase commands are start, stop, pause and resume 
    // Start - start mixing  
    // Stop - stop mixing
    // Pause - stop mixing 
    // Resume - start mixing
    // real states of phase are writed into states in phase structure
    IF MixingPhase.State.ManCtrl THEN
        IF MixingPhase.Cmd.StartMan THEN
            MixingPhase.State.Done := FALSE;
            IF MixingPhase.State.Idle THEN
                MixingPhase.ElapsedTimeSec := 0;
                MixingPhase.State.Idle     := FALSE;
                MixingPhase.State.Paused   := FALSE;
                MixingPhase.State.Running  := TRUE;
            END_IF;
        END_IF;

        IF MixingPhase.Cmd.PauseMan THEN
            MixingPhase.State.Done := FALSE;
            IF MixingPhase.State.Running THEN
                MixingPhase.State.Running := FALSE;
                MixingPhase.State.Idle    := FALSE;
                MixingPhase.State.Paused  := TRUE;
            END_IF;
        END_IF;

        IF MixingPhase.Cmd.ResumeMan THEN
            MixingPhase.State.Done := FALSE;
            IF MixingPhase.State.Paused THEN
                MixingPhase.State.Paused  := FALSE;
                MixingPhase.State.Idle    := FALSE;
                MixingPhase.State.Running := TRUE;
            END_IF;
        END_IF;

        IF MixingPhase.Cmd.StopMan THEN
            MixingPhase.State.Done     := FALSE;
            MixingPhase.State.Running  := FALSE;
            MixingPhase.State.Paused   := FALSE;
            MixingPhase.State.Idle     := TRUE;
            MixingPhase.ElapsedTimeSec := 0;
        END_IF;
    END_IF;

    MixingPhase.Cmd.StartMan  := FALSE;
    MixingPhase.Cmd.StopMan   := FALSE;
    MixingPhase.Cmd.PauseMan  := FALSE;
    MixingPhase.Cmd.ResumeMan := FALSE;
{endregion}

{region "AutCtrl"}
    // if request to run in automatic mode -> set auto request to mixing to 1, if not request to mixing is 0
    // commands should be sets to false after their processing
    IF MixingPhase.State.AutCtrl THEN
        IF MixingPhase.Cmd.StartAut THEN
            MixingPhase.State.Done := FALSE;
            IF MixingPhase.State.Idle THEN
                MixingPhase.ElapsedTimeSec := 0;
                MixingPhase.State.Idle     := FALSE;
                MixingPhase.State.Paused   := FALSE;
                MixingPhase.State.Running  := TRUE;
            END_IF;
        END_IF;

        IF MixingPhase.Cmd.StopAut THEN
            MixingPhase.State.Done     := FALSE;
            MixingPhase.State.Running  := FALSE;
            MixingPhase.State.Paused   := FALSE;
            MixingPhase.State.Idle     := TRUE;
            MixingPhase.ElapsedTimeSec := 0;
        END_IF;
    END_IF;

    MixingPhase.Cmd.StartAut := FALSE;
    MixingPhase.Cmd.StopAut  := FALSE;
{endregion}

{region "Done"}
    // every phase should have finish condition - mixing phase - if time of runnig is bigger or same as requested
    // after that done state should be setted to 1
    secImpTrig(CLK := iSecImp);

    IF MixingPhase.State.Running THEN
        IF secImpTrig.Q THEN
            MixingPhase.ElapsedTimeSec := MixingPhase.ElapsedTimeSec + 1;
        END_IF;

        IF MixingPhase.ElapsedTimeSec >= MixingPhase.ParamTimeSec THEN
            MixingPhase.State.Running  := FALSE;
            MixingPhase.State.Paused   := FALSE;
            MixingPhase.State.Idle     := TRUE;
            MixingPhase.State.Done     := TRUE;
            MixingPhase.ElapsedTimeSec := 0;
        END_IF;
    ELSIF MixingPhase.State.Idle THEN
        MixingPhase.ElapsedTimeSec := 0;
    END_IF;

    IF MixingPhase.Cmd.ResetDone THEN
        MixingPhase.State.Done    := FALSE;
        MixingPhase.Cmd.ResetDone := FALSE;
    END_IF;
{endregion}

{region "States"}
    //Command mixer in cases of states
    IF MixingPhase.State.Running THEN
        MixerEng.Cmd.Req2RunAutCtrl := TRUE;
    ELSE
        MixerEng.Cmd.Req2RunAutCtrl := FALSE;
    END_IF;
{endregion}


// delault state of phase - if not any state sets state to idle
IF NOT MixingPhase.State.Idle AND NOT MixingPhase.State.Paused AND NOT MixingPhase.State.Running THEN
    MixingPhase.State.Idle := 1;
END_IF;


// write binary states into int value for visualization
IF MixingPhase.State.Idle THEN
    MixingPhase.State.StateInt := Global.PhIdle;
ELSIF MixingPhase.State.Running THEN
    MixingPhase.State.StateInt := Global.PhRunning;
ELSE
    MixingPhase.State.StateInt := Global.PhPause;
END_IF;

doEnabled := diEnabled;

END_FUNCTION_BLOCK

// ---- POUs/Draining.TcPOU
FUNCTION_BLOCK Draining
VAR_INPUT
	diEnabled : BOOL;
END_VAR
VAR_OUTPUT
	doEnabled : BOOL;
END_VAR
VAR_IN_OUT
	DrainingPhase : TPhaseDraining;
	DrainingValve : TValve;
END_VAR
VAR
END_VAR

// Synchronizace aktualni hladiny vody (v FB_Tank je RawToEng_1 napojen do Filling.WaterLevel)
DrainingPhase.WaterLevel := Global.Tank1.Filling.WaterLevel;

{region "Aut/Man"}
    // switching state of engine - automatic or manual control (default state is manual)
    IF DrainingPhase.Cmd.ManCtrl THEN
        DrainingPhase.State.ManCtrl := TRUE;
        DrainingPhase.State.AutCtrl := FALSE;
    ELSIF DrainingPhase.Cmd.AutCtrl THEN
        DrainingPhase.State.ManCtrl := FALSE;
        DrainingPhase.State.AutCtrl := TRUE;
    END_IF;

    IF (NOT DrainingPhase.State.ManCtrl) AND (NOT DrainingPhase.State.AutCtrl) THEN
        DrainingPhase.State.ManCtrl := TRUE;
        DrainingPhase.State.AutCtrl := FALSE;
    END_IF;

    DrainingPhase.Cmd.ManCtrl := FALSE;
    DrainingPhase.Cmd.AutCtrl := FALSE;
{endregion}

{region "ManCtrl"}
    // processing manual actions - if command is processed, it is sets to FALSE even if can't be processed
    // Phase commands are start, stop, pause and resume 
    // Start - open draining valve 
    // Stop - close draining valve
    // Pause - close draining valve
    // Resume - open draining valve
    // real states of phase are writed into states in phase structure
    IF DrainingPhase.State.ManCtrl THEN
        IF DrainingPhase.Cmd.StartMan THEN
            DrainingPhase.State.Done := FALSE;
            IF DrainingPhase.State.Idle THEN
                DrainingPhase.State.Idle    := FALSE;
                DrainingPhase.State.Paused  := FALSE;
                DrainingPhase.State.Running := TRUE;
            END_IF;
        END_IF;

        IF DrainingPhase.Cmd.PauseMan THEN
            DrainingPhase.State.Done := FALSE;
            IF DrainingPhase.State.Running THEN
                DrainingPhase.State.Running := FALSE;
                DrainingPhase.State.Idle    := FALSE;
                DrainingPhase.State.Paused  := TRUE;
            END_IF;
        END_IF;

        IF DrainingPhase.Cmd.ResumeMan THEN
            DrainingPhase.State.Done := FALSE;
            IF DrainingPhase.State.Paused THEN
                DrainingPhase.State.Paused  := FALSE;
                DrainingPhase.State.Idle    := FALSE;
                DrainingPhase.State.Running := TRUE;
            END_IF;
        END_IF;

        IF DrainingPhase.Cmd.StopMan THEN
            DrainingPhase.State.Done    := FALSE;
            DrainingPhase.State.Running := FALSE;
            DrainingPhase.State.Paused  := FALSE;
            DrainingPhase.State.Idle    := TRUE;
        END_IF;
    END_IF;

    DrainingPhase.Cmd.StartMan  := FALSE;
    DrainingPhase.Cmd.StopMan   := FALSE;
    DrainingPhase.Cmd.PauseMan  := FALSE;
    DrainingPhase.Cmd.ResumeMan := FALSE;
{endregion}

{region "AutCtrl"}
    //if request to run in automatic mode -> set auto request to open of filling valve to 1 and close to 0, if not open 0 close 1
    // commands should be sets to false after their processing
    IF DrainingPhase.State.AutCtrl THEN
        IF DrainingPhase.Cmd.StartAut THEN
            DrainingPhase.State.Done := FALSE;
            IF DrainingPhase.State.Idle THEN
                DrainingPhase.State.Idle    := FALSE;
                DrainingPhase.State.Paused  := FALSE;
                DrainingPhase.State.Running := TRUE;
            END_IF;
        END_IF;

        IF DrainingPhase.Cmd.StopAut THEN
            DrainingPhase.State.Done    := FALSE;
            DrainingPhase.State.Running := FALSE;
            DrainingPhase.State.Paused  := FALSE;
            DrainingPhase.State.Idle    := TRUE;
        END_IF;
    END_IF;

    DrainingPhase.Cmd.StartAut := FALSE;
    DrainingPhase.Cmd.StopAut  := FALSE;
{endregion}
{region "Done"}
    //every phase should have finish condition - draining phase - if water level is below requested level
    //after that done state should be setted to 1
    IF DrainingPhase.State.Running THEN
        IF DrainingPhase.WaterLevel <= DrainingPhase.ParamDrainLevel THEN
            DrainingPhase.State.Running := FALSE;
            DrainingPhase.State.Paused  := FALSE;
            DrainingPhase.State.Idle    := TRUE;
            DrainingPhase.State.Done    := TRUE;
        END_IF;
    END_IF;

    IF DrainingPhase.Cmd.ResetDone THEN
        DrainingPhase.State.Done    := FALSE;
        DrainingPhase.Cmd.ResetDone := FALSE;
    END_IF;
{endregion}

{region "States"} 
    //Command valve in cases of states
    IF DrainingPhase.State.Running THEN
        DrainingValve.Cmd.Req2OpenAut  := TRUE;
        DrainingValve.Cmd.Req2CloseAut := FALSE;
    ELSE
        DrainingValve.Cmd.Req2OpenAut  := FALSE;
        DrainingValve.Cmd.Req2CloseAut := TRUE;
    END_IF;
{endregion}

// delault state of phase - if not any state sets state to idle
IF (NOT DrainingPhase.State.Idle) AND (NOT DrainingPhase.State.Paused) AND (NOT DrainingPhase.State.Running) THEN
    DrainingPhase.State.Idle := 1;
END_IF;

// write binary states into int value for visualization
IF DrainingPhase.State.Idle THEN
    DrainingPhase.State.StateInt := Global.PhIdle;
ELSIF DrainingPhase.State.Running THEN
    DrainingPhase.State.StateInt := Global.PhRunning;
ELSE
    DrainingPhase.State.StateInt := Global.PhPause;
END_IF;

//Ponechte pro moznost retezeni volani bloku v LAD
doEnabled := diEnabled;

END_FUNCTION_BLOCK

// ---- POUs/Heating.TcPOU
FUNCTION_BLOCK Heating
VAR_INPUT
	diEnabled : BOOL;
	iSecImp : BOOL;
END_VAR
VAR_OUTPUT
	doEnabled : BOOL;
END_VAR
VAR_IN_OUT
	HeatingPhase : TPhaseHeating;
	Heater : THeater;
END_VAR
VAR
	pidParameters : ST_CTRL_PID_PARAMS;
	secImpTrig : R_TRIG;
END_VAR

{region "Aut/Man"}
    // switching state of engine - automatic or manual control (default state is manual)
    IF HeatingPhase.Cmd.ManCtrl THEN
        HeatingPhase.State.ManCtrl := TRUE;
        HeatingPhase.State.AutCtrl := FALSE;
    ELSIF HeatingPhase.Cmd.AutCtrl THEN
        HeatingPhase.State.ManCtrl := FALSE;
        HeatingPhase.State.AutCtrl := TRUE;
    END_IF;

    IF (NOT HeatingPhase.State.ManCtrl) AND (NOT HeatingPhase.State.AutCtrl) THEN
        HeatingPhase.State.ManCtrl := TRUE;
        HeatingPhase.State.AutCtrl := FALSE;
    END_IF;

    HeatingPhase.Cmd.ManCtrl := FALSE;
    HeatingPhase.Cmd.AutCtrl := FALSE;
{endregion}

{region "ManCtrl"}
    // processing manual actions - if command is processed, it is sets to FALSE even if can't be processed
    // real states of phase are writed into states in phase structure
    IF HeatingPhase.State.ManCtrl THEN
        IF HeatingPhase.Cmd.StartMan THEN
            HeatingPhase.State.Done := FALSE;
            IF HeatingPhase.State.Idle THEN
                HeatingPhase.fTime         := 0;
                HeatingPhase.State.Idle    := FALSE;
                HeatingPhase.State.Paused  := FALSE;
                HeatingPhase.State.Running := TRUE;
            END_IF;
        END_IF;

        IF HeatingPhase.Cmd.PauseMan THEN
            HeatingPhase.State.Done := FALSE;
            IF HeatingPhase.State.Running THEN
                HeatingPhase.State.Running := FALSE;
                HeatingPhase.State.Idle    := FALSE;
                HeatingPhase.State.Paused  := TRUE;
            END_IF;
        END_IF;

        IF HeatingPhase.Cmd.ResumeMan THEN
            HeatingPhase.State.Done := FALSE;
            IF HeatingPhase.State.Paused THEN
                HeatingPhase.State.Paused  := FALSE;
                HeatingPhase.State.Idle    := FALSE;
                HeatingPhase.State.Running := TRUE;
            END_IF;
        END_IF;

        IF HeatingPhase.Cmd.StopMan THEN
            HeatingPhase.State.Done    := FALSE;
            HeatingPhase.State.Running := FALSE;
            HeatingPhase.State.Paused  := FALSE;
            HeatingPhase.State.Idle    := TRUE;
            HeatingPhase.fTime         := 0;
        END_IF;
    END_IF;

    HeatingPhase.Cmd.StartMan  := FALSE;
    HeatingPhase.Cmd.StopMan   := FALSE;
    HeatingPhase.Cmd.PauseMan  := FALSE;
    HeatingPhase.Cmd.ResumeMan := FALSE;
{endregion}

{region "AutCtrl"}
    // if request to run in automatic mode -> set auto request to heat to 1, if not request to heat 0
    // commands should be sets to false after their processing
    IF HeatingPhase.State.AutCtrl THEN
        IF HeatingPhase.Cmd.StartAut THEN
            HeatingPhase.State.Done := FALSE;
            IF HeatingPhase.State.Idle THEN
                HeatingPhase.fTime         := 0;
                HeatingPhase.State.Idle    := FALSE;
                HeatingPhase.State.Paused  := FALSE;
                HeatingPhase.State.Running := TRUE;
            END_IF;
        END_IF;

        IF HeatingPhase.Cmd.StopAut THEN
            HeatingPhase.State.Done    := FALSE;
            HeatingPhase.State.Running := FALSE;
            HeatingPhase.State.Paused  := FALSE;
            HeatingPhase.State.Idle    := TRUE;
            HeatingPhase.fTime         := 0;
        END_IF;
    END_IF;

    HeatingPhase.Cmd.StartAut := FALSE;
    HeatingPhase.Cmd.StopAut  := FALSE;
{endregion}

{region "Done"}
    //every phase should have finish condition - heating phase - if water temp is on requested value for 10 seconds with 1°C hysteresis
    //after that done state should be setted to 1
    secImpTrig(CLK := iSecImp);

    IF HeatingPhase.State.Running THEN
        IF (HeatingPhase.WaterTemp >= (HeatingPhase.ParamReqTemp - 1.0)) AND (HeatingPhase.WaterTemp <= (HeatingPhase.ParamReqTemp + 1.0)) THEN
            IF secImpTrig.Q THEN
                HeatingPhase.fTime := HeatingPhase.fTime + 1;
            END_IF;
        ELSE
            HeatingPhase.fTime := 0;
        END_IF;

        IF HeatingPhase.fTime >= 1 THEN				/// TADY MA BYT 10
            HeatingPhase.State.Running := FALSE;
            HeatingPhase.State.Paused  := FALSE;
            HeatingPhase.State.Idle    := TRUE;
            HeatingPhase.State.Done    := TRUE;
            HeatingPhase.fTime         := 0;
        END_IF;
    ELSE
        HeatingPhase.fTime := 0;
    END_IF;

    // command reset done resets done state and than resets command
    IF HeatingPhase.Cmd.ResetDone THEN
        HeatingPhase.State.Done    := FALSE;
        HeatingPhase.Cmd.ResetDone := FALSE;
    END_IF;
{endregion}

{region "States"}
    //Command valve in cases of states
    // Running - start heating  
    // Idle - stop heating
    // Pause - stop heating (alternative is hold actual temp)
    IF HeatingPhase.State.Running THEN
        Heater.ParamHeatingSetPointAutomat := HeatingPhase.ParamReqTemp;
        Heater.Cmd.Req2RunAutCtrl := TRUE;
    ELSE
        Heater.Cmd.Req2RunAutCtrl := FALSE;
    END_IF;
{endregion}

// delault state of phase - if not any state sets state to idle
IF NOT HeatingPhase.State.Idle AND NOT HeatingPhase.State.Paused AND NOT HeatingPhase.State.Running THEN
    HeatingPhase.State.Idle := 1;
END_IF;

// write binary states into int value for visualization
IF HeatingPhase.State.Idle THEN
    HeatingPhase.State.Stateint := Global.PhIdle;
ELSIF HeatingPhase.State.Running THEN
    HeatingPhase.State.Stateint := Global.PhRunning;
ELSE
    HeatingPhase.State.Stateint := Global.PhPause;
END_IF;

doEnabled := diEnabled;

END_FUNCTION_BLOCK

// ---- POUs/Misc/RawToEng.TcPOU
FUNCTION_BLOCK RawToEng
VAR_INPUT
	iEnabled : BOOL;
	wRawValue : WORD;
	AnalogConversion : TAnalogConversion;
END_VAR
VAR_OUTPUT
	oEnabled : BOOL;
	fScaledValue : REAL;
END_VAR
VAR
END_VAR

//Prepocet z wRawValue (z procesu po ModbusTCP) na fScaledValue (do PLC) podle parametru v AnalogConversion.

//Filtrace hodnoty: odfiltrovani skokoveho kmitani z minimalniho rozsahu na maximalni hodnotu >= 27648 (podteceni sumu u nuly v simulatoru)
IF wRawValue >= AnalogConversion.TransducerHiLevel THEN 
	IF fScaledValue < ((AnalogConversion.ScaledValHiLevel + AnalogConversion.ScaledValLoLevel) / 2.0) THEN
		wRawValue := AnalogConversion.TransducerLoLevel;
	ELSE
		wRawValue := AnalogConversion.TransducerHiLevel;
	END_IF;
END_IF;

fScaledValue := (AnalogConversion.ScaledValHiLevel - AnalogConversion.ScaledValLoLevel) * WORD_TO_REAL(wRawValue - AnalogConversion.TransducerLoLevel) / UINT_TO_REAL(AnalogConversion.TransducerHiLevel - AnalogConversion.TransducerLoLevel) + AnalogConversion.ScaledValLoLevel;
oEnabled := iEnabled;

END_FUNCTION_BLOCK

// ---- POUs/Misc/EngToRaw.TcPOU
FUNCTION_BLOCK EngToRaw
VAR_INPUT
	iEnabled : BOOL;
	fScaledValue : REAL;
	AnalogConversion : TAnalogConversion;
END_VAR
VAR_OUTPUT
	oEnabled : BOOL;
	wRawValue : WORD;
END_VAR
VAR
END_VAR

//Prepocet z fScaledValue (z PLC) na wRawValue (do procesu po ModbusTCP) podle parametru v AnalogConversion.
IF fScaledValue <= AnalogConversion.ScaledValLoLevel THEN
	wRawValue := UINT_TO_WORD(AnalogConversion.TransducerLoLevel);
ELSIF fScaledValue >= AnalogConversion.ScaledValHiLevel THEN
	wRawValue := UINT_TO_WORD(AnalogConversion.TransducerHiLevel);
ELSE
	wRawValue := REAL_TO_WORD(UINT_TO_REAL(AnalogConversion.TransducerHiLevel - AnalogConversion.TransducerLoLevel) * (fScaledValue - AnalogConversion.ScaledValLoLevel) / (AnalogConversion.ScaledValHiLevel - AnalogConversion.ScaledValLoLevel) + UINT_TO_REAL(AnalogConversion.TransducerLoLevel));
END_IF;
oEnabled := iEnabled;

END_FUNCTION_BLOCK

// ---- POUs/MAIN.TcPOU
PROGRAM MAIN
VAR
	// --- PŘEPÍNAČ PŘÍMÉHO RUČNÍHO TESTOVÁNÍ SIMULÁTORU ---
	// FALSE = výstupy řídí FB_Tank_1 v Main_Batch (standardní provoz)
	// TRUE  = výstupy řídí přímo proměnné bTest_* níže (pouze když je zakomentovaný Main_Batch)
	bTest_ManualOverride  : BOOL := FALSE;
	test_prom : BOOL;
	// --- RUČNÍ TESTOVACÍ OVLÁDÁNÍ AKČNÍCH ČLENŮ (Zápis do simulátoru) ---
	bTest_FillValve_Open  : BOOL := FALSE; // TRUE = otevírá napouštěcí ventil, FALSE = aktivně zavírá
	bTest_DrainValve_Open : BOOL := FALSE; // TRUE = otevírá vypouštěcí ventil, FALSE = aktivně zavírá
	bTest_Mixer           : BOOL := FALSE; // TRUE = zapne míchadlo
	bTest_Heating         : BOOL := FALSE; // TRUE = povolí topení a pošle wTest_HeatingPower
	wTest_HeatingPower    : WORD := 15000; // Požadovaný výkon topení (0..27648 odpovídá 0..100 %)

	// --- ČTENÍ STAVŮ ZE SIMULÁTORU (Pro přehled v Online režimu) ---
	// Napouštěcí ventil (koncové dorazy a porucha)
	bStat_FillValve_IsOpen   : BOOL;
	bStat_FillValve_IsClosed : BOOL;
	bStat_FillValve_Error    : BOOL;

	// Vypouštěcí ventil (koncové dorazy a porucha)
	bStat_DrainValve_IsOpen   : BOOL;
	bStat_DrainValve_IsClosed : BOOL;
	bStat_DrainValve_Error    : BOOL;

	// Míchadlo (zpětná vazba chodu a porucha)
	bStat_Mixer_IsRunning : BOOL;
	bStat_Mixer_Error     : BOOL;

	// Spojité snímače (surové hodnoty 0..27648 i přepočet na m a °C)
	wStat_WaterLevel_Raw : WORD;
	fStat_WaterLevel_m   : REAL; // Přepočtená hladina (0.0 .. 2.0 m)
	wStat_WaterTemp_Raw  : WORD;
	fStat_WaterTemp_C    : REAL; // Přepočtená teplota (0.0 .. 100.0 °C)
END_VAR

// Generování hodinového impulzu s periodou 1 s (MAIN běží v PlcTask500ms s periodou 500 ms)
Global.secImp := NOT(Global.secImp);

// ============================================================================
// 1. ZÁPIS TESTOVACÍCH POVELŮ DO SIMULÁTORU (pouze pokud je bTest_ManualOverride = TRUE)
//    Při standardním běhu přes FB_Tank_1 v Main_Batch musí být bTest_ManualOverride = FALSE!
// ============================================================================
IF bTest_ManualOverride THEN
	// Napouštěcí ventil (v maup.NET drží bez povelu poslední stav -> při FALSE aktivně zavíráme)
	IF bTest_FillValve_Open THEN
		Global.doValveFillOpen  := TRUE;
		Global.doValveFillClose := FALSE;
	ELSE
		Global.doValveFillOpen  := FALSE;
		Global.doValveFillClose := TRUE;
	END_IF;

	// Vypouštěcí ventil (při FALSE aktivně zavíráme)
	IF bTest_DrainValve_Open THEN
		Global.doValveDrainOpen  := TRUE;
		Global.doValveDrainClose := FALSE;
	ELSE
		Global.doValveDrainOpen  := FALSE;
		Global.doValveDrainClose := TRUE;
	END_IF;

	// Míchadlo
	Global.doMixerStart := bTest_Mixer;

	// Ohřev (odblokování topení + výkon do holding registru)
	Global.doHeatingEnable := bTest_Heating;
	IF bTest_Heating THEN
		Global.aoReqPowerOfHeating := wTest_HeatingPower;
	ELSE
		Global.aoReqPowerOfHeating := 0;
	END_IF;
ELSE
	test_prom :=false;
END_IF;

// ============================================================================
// 2. ČTENÍ STAVŮ A SENZORŮ ZE SIMULÁTORU (z Global.di* a Global.ai*)
//    (Běží neustále – pouze čte hodnoty pro rychlou diagnostiku v Online režimu)
// ============================================================================

// Napouštěcí ventil
bStat_FillValve_IsOpen   := Global.diValveFillOpen;
bStat_FillValve_IsClosed := Global.diValveFillClose;
bStat_FillValve_Error    := Global.diValveFillError;

// Vypouštěcí ventil
bStat_DrainValve_IsOpen   := Global.diValveDrainOpen;
bStat_DrainValve_IsClosed := Global.diValveDrainClose;
bStat_DrainValve_Error    := Global.diValveDrainError;

// Míchadlo
bStat_Mixer_IsRunning := Global.diMixerRun;
bStat_Mixer_Error     := Global.diMixerError;

// Analogové hodnoty (surové 0..27648 + orientační přepočet na fyzikální jednotky)
wStat_WaterLevel_Raw := Global.aiWaterLevel;
fStat_WaterLevel_m   := WORD_TO_REAL(Global.aiWaterLevel) * 2.0 / 27648.0;

wStat_WaterTemp_Raw  := Global.aiWaterTemp;
fStat_WaterTemp_C    := WORD_TO_REAL(Global.aiWaterTemp) * 100.0 / 27648.0;

// Volani hlavniho davkoveho automatu (kap. 10.4)
Test();

END_PROGRAM

// ---- POUs/Test.TcPOU
PROGRAM Test
VAR
	State             : INT := 0;       // 0=Idle, 10=Init/Aut, 20..25=Filling, 30..35=Mix+Heat, 40..45=Draining, 50=NextBatch
	bStartBatch       : BOOL := FALSE;  // Prikaz pro spusteni davkove vyroby
	bStopBatch        : BOOL := FALSE;  // Prikaz pro okamzite zastaveni vyroby
	bRunning          : BOOL := FALSE;  // Signalizace, ze automat prave bezi
	nTargetBatches    : INT := 1;       // Pozadovany pocet davek
	nCompletedBatches : INT := 0;       // Pocet jiz vyrobenych davek
	bInitDone         : BOOL := FALSE;  // Jednorazova inicializace vychozich parametru receptury
END_VAR

// Jednorazova inicializace vychozich parametru receptury po startu PLC (pokud jsou 0)
IF NOT bInitDone THEN
	IF Global.Tank1.Filling.ParamFillLevel <= 0.0 THEN
		Global.Tank1.Filling.ParamFillLevel := 1.0;
	END_IF;
	IF Global.Tank1.Draining.ParamDrainLevel <= 0.0 THEN
		Global.Tank1.Draining.ParamDrainLevel := 0.2;
	END_IF;
	IF Global.Tank1.Mixing.ParamTimeSec <= 0 THEN
		Global.Tank1.Mixing.ParamTimeSec := 10;
	END_IF;
	IF Global.Tank1.Heating.ParamReqTemp <= 0.0 THEN
		Global.Tank1.Heating.ParamReqTemp := 40.0;
	END_IF;
	bInitDone := TRUE;
END_IF;

// Okamzite zastaveni automatu pri prikazu Stop nebo pri chybe GlobalError
IF bStopBatch OR (bRunning AND Global.Tank1.GlobalError) THEN
	Global.Tank1.Filling.Cmd.StopAut  := TRUE;
	Global.Tank1.Draining.Cmd.StopAut := TRUE;
	Global.Tank1.Mixing.Cmd.StopAut   := TRUE;
	Global.Tank1.Heating.Cmd.StopAut  := TRUE;
	bRunning   := FALSE;
	State      := 0;
	bStopBatch := FALSE;
END_IF;

CASE State OF
	0: // Idle - cekani na prikaz Start Batch
		bRunning := FALSE;
		IF bStartBatch THEN
			IF nTargetBatches < 1 THEN
				nTargetBatches := 1;
			END_IF;
			nCompletedBatches := 0;
			bRunning := TRUE;
			State    := 10;
		END_IF;

	10: // Prepne vsechny akcni cleny i faze do AUT a vymaze stare priznaky Done
		Global.Tank1.ValveFilling.Cmd.AutCtrl  := TRUE;
		Global.Tank1.ValveDraining.Cmd.AutCtrl := TRUE;
		Global.Tank1.Mixer.Cmd.AutCtrl         := TRUE;
		Global.Tank1.Heater.Cmd.AutCtrl        := TRUE;

		Global.Tank1.Filling.Cmd.AutCtrl   := TRUE;
		Global.Tank1.Draining.Cmd.AutCtrl  := TRUE;
		Global.Tank1.Mixing.Cmd.AutCtrl    := TRUE;
		Global.Tank1.Heating.Cmd.AutCtrl   := TRUE;

		Global.Tank1.Filling.Cmd.ResetDone  := TRUE;
		Global.Tank1.Draining.Cmd.ResetDone := TRUE;
		Global.Tank1.Mixing.Cmd.ResetDone   := TRUE;
		Global.Tank1.Heating.Cmd.ResetDone  := TRUE;

		State := 20;

	20: // Spusteni faze napousteni (Filling)
		IF Global.Tank1.Filling.State.AutCtrl THEN
			Global.Tank1.Filling.Cmd.StartAut := TRUE;
			State := 25;
		END_IF;

	25: // Cekani na dokonceni napousteni
		IF Global.Tank1.Filling.State.Done THEN
			Global.Tank1.Filling.Cmd.ResetDone := TRUE;
			State := 30;
		END_IF;

	30: // Spusteni soubeznych fazi michani a ohrevu (Mixing + Heating)
		IF Global.Tank1.Mixing.State.AutCtrl AND Global.Tank1.Heating.State.AutCtrl THEN
			Global.Tank1.Mixing.Cmd.StartAut  := TRUE;
			Global.Tank1.Heating.Cmd.StartAut := TRUE;
			State := 35;
		END_IF;

	35: // Cekani na dokonceni michani I ohrevu
		IF Global.Tank1.Mixing.State.Done AND Global.Tank1.Heating.State.Done THEN
			Global.Tank1.Mixing.Cmd.ResetDone  := TRUE;
			Global.Tank1.Heating.Cmd.ResetDone := TRUE;
			State := 40;
		END_IF;

	40: // Spusteni faze vypousteni (Draining)
		IF Global.Tank1.Draining.State.AutCtrl THEN
			Global.Tank1.Draining.Cmd.StartAut := TRUE;
			State := 45;
		END_IF;

	45: // Cekani na dokonceni vypousteni
		IF Global.Tank1.Draining.State.Done THEN
			Global.Tank1.Draining.Cmd.ResetDone := TRUE;
			State := 50;
		END_IF;

	50: // Vyhodnoceni poctu vyrobenych davek
		nCompletedBatches := nCompletedBatches + 1;
		IF nCompletedBatches < nTargetBatches THEN
			State := 10; // Dalsi davka
		ELSE
			bRunning := FALSE;
			State    := 0;  // Hotovo
		END_IF;
END_CASE;

bStartBatch := FALSE;

END_PROGRAM

// ---- GlobalTextList.TcGTLO
TEXTLIST GlobalTextList
  815 = 'ABC'
  406 = 'AUT'
  473 = 'Checkbox'
  70 = 'Close'
  25 = 'Closed'
  201 = 'Filling Valve'
  560 = 'MAN'
  604 = 'Open'
  687 = 'Opened'
  98 = 'Res. SUF'
  256 = 'SUF'
  202 = 'Draining Valve'
  203 = 'Mixer'
  204 = 'Heater'
  205 = 'Stop'
  206 = 'Turn On'
  207 = 'Turn Off'
  208 = 'Run'
  209 = 'Err'
  210 = 'RT: %d s'
  211 = 'SetRT: %d'
  212 = 'Man Pwr: %.1f %%'
  213 = 'Aut Set: %.1f C'
  214 = 'Out'
  215 = '%.0f %%'
  216 = 'Level: %.2f m'
  217 = 'Temp: %.1f C'
  218 = 'Global Err'
  219 = 'Phase: Filling'
  220 = 'Phase: Draining'
  221 = 'Phase: Mixing'
  222 = 'Phase: Heating'
  223 = 'Idle'
  224 = 'Pause'
  225 = 'Done'
  226 = 'Start'
  227 = 'Resume'
  228 = 'Res.Done'
  229 = 'Fill Lvl: %.2f m'
  230 = 'Drain Lvl: %.2f m'
  231 = 'Mix Time: %d s'
  232 = 'Req Temp: %.1f C'
  233 = 'Act: %.2f m'
  234 = 'Elap: %d s'
  235 = 'Hold: %d s'
  236 = 'Batch Automat (Test)'
  237 = 'Start Batch'
  238 = 'Stop Batch'
  239 = 'Batches: %d'
  240 = 'Done: %d'
  241 = 'Step: %d'
END_TEXTLIST

// ---- VISUs/Visualization.TcVIS
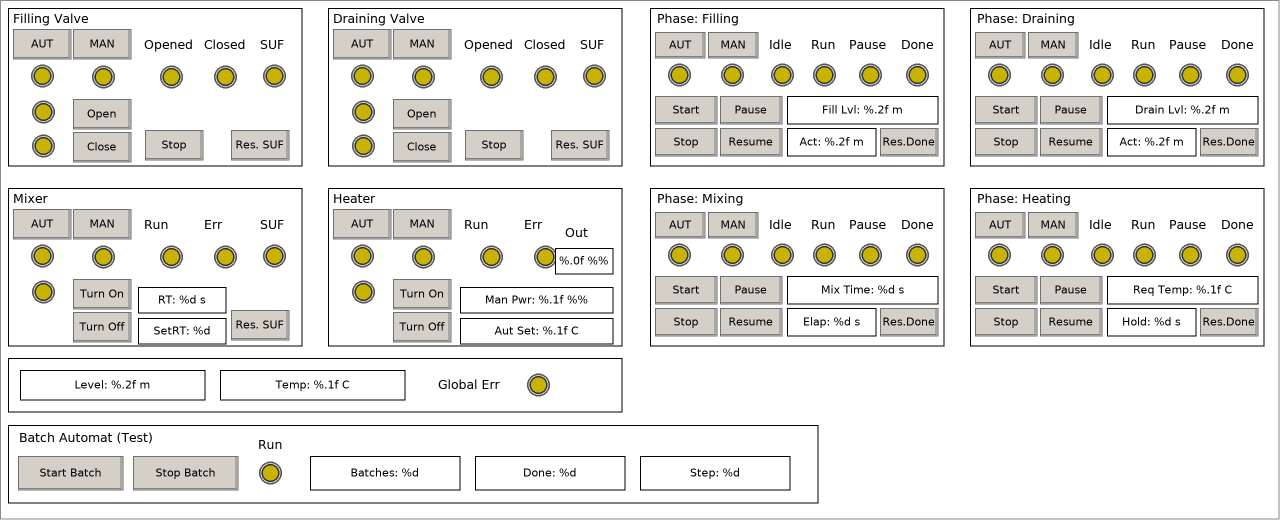
VISUALIZATION Visualization  // 1280x520
    Rectangle (8,8 294x158)
    Button (13,29 58x30), "AUT"
        OnMouseClick: toggle Global.Tank1.ValveFilling.Cmd.AutCtrl
    Button (73,29 58x30), "MAN"
        OnMouseClick: toggle Global.Tank1.ValveFilling.Cmd.ManCtrl
    Label (10,10 96x18), "Filling Valve"
    Button (73,99 58x30), "Open"
        OnMouseClick: toggle Global.Tank1.ValveFilling.Cmd.OpenMan
    Button (73,132 58x30), "Close"
        OnMouseClick: toggle Global.Tank1.ValveFilling.Cmd.CloseMan
    Lamp1 (29,63 27x26), variable: Global.Tank1.ValveFilling.State.AutCtrl, style: Lamp-Lamp1-Yellow
    Lamp1 (90,64 27x26), variable: Global.Tank1.ValveFilling.State.ManCtrl, style: Lamp-Lamp1-Yellow
    Lamp1 (158,64 27x26), variable: Global.Tank1.ValveFilling.State.Open, style: Lamp-Lamp1-Yellow
    Lamp1 (212,64 27x26), variable: Global.Tank1.ValveFilling.State.Closed, style: Lamp-Lamp1-Yellow
    Lamp1 (261,63 27x26), variable: Global.Tank1.ValveFilling.State.StartupFail, style: Lamp-Lamp1-Yellow
    Button (231,130 58x30), "Res. SUF"
        OnMouseClick: toggle Global.Tank1.ValveFilling.Cmd.ResetSUF
    Label (141,36 53x18), "Opened"
    Label (201,36 53x18), "Closed"
    Label (257,36 33x18), "SUF"
    Lamp1 (30,99 27x26), variable: Global.Tank1.ValveFilling.State.OpenOut, style: Lamp-Lamp1-Yellow
    Lamp1 (30,133 27x26), variable: Global.Tank1.ValveFilling.State.CloseOut, style: Lamp-Lamp1-Yellow
    Button (145,130 58x30), "Stop"
        OnMouseClick: toggle Global.Tank1.ValveFilling.Cmd.StopMan
    Rectangle (328,8 294x158)
    Button (333,29 58x30), "AUT"
        OnMouseClick: toggle Global.Tank1.ValveDraining.Cmd.AutCtrl
    Button (393,29 58x30), "MAN"
        OnMouseClick: toggle Global.Tank1.ValveDraining.Cmd.ManCtrl
    Label (330,10 120x18), "Draining Valve"
    Button (393,99 58x30), "Open"
        OnMouseClick: toggle Global.Tank1.ValveDraining.Cmd.OpenMan
    Button (393,132 58x30), "Close"
        OnMouseClick: toggle Global.Tank1.ValveDraining.Cmd.CloseMan
    Lamp1 (349,63 27x26), variable: Global.Tank1.ValveDraining.State.AutCtrl, style: Lamp-Lamp1-Yellow
    Lamp1 (410,64 27x26), variable: Global.Tank1.ValveDraining.State.ManCtrl, style: Lamp-Lamp1-Yellow
    Lamp1 (478,64 27x26), variable: Global.Tank1.ValveDraining.State.Open, style: Lamp-Lamp1-Yellow
    Lamp1 (532,64 27x26), variable: Global.Tank1.ValveDraining.State.Closed, style: Lamp-Lamp1-Yellow
    Lamp1 (581,63 27x26), variable: Global.Tank1.ValveDraining.State.StartupFail, style: Lamp-Lamp1-Yellow
    Button (551,130 58x30), "Res. SUF"
        OnMouseClick: toggle Global.Tank1.ValveDraining.Cmd.ResetSUF
    Label (461,36 53x18), "Opened"
    Label (521,36 53x18), "Closed"
    Label (577,36 33x18), "SUF"
    Lamp1 (350,99 27x26), variable: Global.Tank1.ValveDraining.State.OpenOut, style: Lamp-Lamp1-Yellow
    Lamp1 (350,133 27x26), variable: Global.Tank1.ValveDraining.State.CloseOut, style: Lamp-Lamp1-Yellow
    Button (465,130 58x30), "Stop"
        OnMouseClick: toggle Global.Tank1.ValveDraining.Cmd.StopMan
    Rectangle (8,188 294x158)
    Button (13,209 58x30), "AUT"
        OnMouseClick: toggle Global.Tank1.Mixer.Cmd.AutCtrl
    Button (73,209 58x30), "MAN"
        OnMouseClick: toggle Global.Tank1.Mixer.Cmd.ManCtrl
    Label (10,190 96x18), "Mixer"
    Button (73,279 58x30), "Turn On"
        OnMouseClick: toggle Global.Tank1.Mixer.Cmd.TurnOnMan
    Button (73,312 58x30), "Turn Off"
        OnMouseClick: toggle Global.Tank1.Mixer.Cmd.TurnOffMan
    Lamp1 (29,243 27x26), variable: Global.Tank1.Mixer.State.AutCtrl, style: Lamp-Lamp1-Yellow
    Lamp1 (90,244 27x26), variable: Global.Tank1.Mixer.State.ManCtrl, style: Lamp-Lamp1-Yellow
    Lamp1 (158,244 27x26), variable: Global.Tank1.Mixer.State.Run, style: Lamp-Lamp1-Yellow
    Lamp1 (212,244 27x26), variable: Global.Tank1.Mixer.State.GenErr, style: Lamp-Lamp1-Yellow
    Lamp1 (261,243 27x26), variable: Global.Tank1.Mixer.State.StartUpFail, style: Lamp-Lamp1-Yellow
    Button (231,310 58x30), "Res. SUF"
        OnMouseClick: toggle Global.Tank1.Mixer.Cmd.ResetSUF
    Label (141,216 53x18), "Run"
    Label (201,216 53x18), "Err"
    Label (257,216 33x18), "SUF"
    Lamp1 (30,279 27x26), variable: Global.Tank1.Mixer.State.RunOut, style: Lamp-Lamp1-Yellow
    Rectangle (328,188 294x158)
    Button (333,209 58x30), "AUT"
        OnMouseClick: toggle Global.Tank1.Heater.Cmd.AutCtrl
    Button (393,209 58x30), "MAN"
        OnMouseClick: toggle Global.Tank1.Heater.Cmd.ManCtrl
    Label (330,190 96x18), "Heater"
    Button (393,279 58x30), "Turn On"
        OnMouseClick: toggle Global.Tank1.Heater.Cmd.TurnOnMan
    Button (393,312 58x30), "Turn Off"
        OnMouseClick: toggle Global.Tank1.Heater.Cmd.TurnOffMan
    Lamp1 (349,243 27x26), variable: Global.Tank1.Heater.State.AutCtrl, style: Lamp-Lamp1-Yellow
    Lamp1 (410,244 27x26), variable: Global.Tank1.Heater.State.ManCtrl, style: Lamp-Lamp1-Yellow
    Lamp1 (478,244 27x26), variable: Global.Tank1.Heater.State.EnableOut, style: Lamp-Lamp1-Yellow
    Lamp1 (532,244 27x26), variable: Global.Tank1.Heater.State.GenErr, style: Lamp-Lamp1-Yellow
    Label (461,216 53x18), "Run"
    Label (521,216 53x18), "Err"
    Lamp1 (350,279 27x26), variable: Global.Tank1.Heater.State.EnableOut, style: Lamp-Lamp1-Yellow
    Rectangle (138,287 88x26), "RT: %d s", text variable: Global.Tank1.Mixer.State.RT
    Rectangle (138,318 88x26), "SetRT: %d", text variable: Global.Tank1.Mixer.Cmd.SetRT
        OnMouseClick: write the text variable via Default
    Label (562,224 45x18), "Out"
    Rectangle (555,248 58x26), "%.0f %%", text variable: Global.Tank1.Heater.State.HeatingOut
    Rectangle (460,287 153x26), "Man Pwr: %.1f %%", text variable: Global.Tank1.Heater.ParamHeatingPowerManual
        OnMouseClick: write the text variable via Default
    Rectangle (460,318 153x26), "Aut Set: %.1f C", text variable: Global.Tank1.Heater.ParamHeatingSetPointAutomat
        OnMouseClick: write the text variable via Default
    Rectangle (8,358 614x54)
    Rectangle (20,370 185x30), "Level: %.2f m", text variable: Global.Tank1.Filling.WaterLevel
    Rectangle (220,370 185x30), "Temp: %.1f C", text variable: Global.Tank1.Heating.WaterTemp
    Label (435,376 85x20), "Global Err"
    Lamp1 (525,372 27x26), variable: Global.Tank1.GlobalError, style: Lamp-Lamp1-Yellow
    Rectangle (650,8 294x158)
    Label (654,10 140x18), "Phase: Filling"
    Button (655,32 50x26), "AUT"
        OnMouseClick: toggle Global.Tank1.Filling.Cmd.AutCtrl
    Button (708,32 50x26), "MAN"
        OnMouseClick: toggle Global.Tank1.Filling.Cmd.ManCtrl
    Label (766,36 38x18), "Idle"
    Label (808,36 38x18), "Run"
    Label (846,36 52x18), "Pause"
    Label (898,36 44x18), "Done"
    Lamp1 (666,62 27x26), variable: Global.Tank1.Filling.State.AutCtrl, style: Lamp-Lamp1-Yellow
    Lamp1 (719,62 27x26), variable: Global.Tank1.Filling.State.ManCtrl, style: Lamp-Lamp1-Yellow
    Lamp1 (769,62 27x26), variable: Global.Tank1.Filling.State.Idle, style: Lamp-Lamp1-Yellow
    Lamp1 (811,62 27x26), variable: Global.Tank1.Filling.State.Running, style: Lamp-Lamp1-Yellow
    Lamp1 (857,62 27x26), variable: Global.Tank1.Filling.State.Paused, style: Lamp-Lamp1-Yellow
    Lamp1 (904,62 27x26), variable: Global.Tank1.Filling.State.Done, style: Lamp-Lamp1-Yellow
    Button (655,96 62x28), "Start"
        OnMouseClick: toggle Global.Tank1.Filling.Cmd.StartMan
    Button (720,96 62x28), "Pause"
        OnMouseClick: toggle Global.Tank1.Filling.Cmd.PauseMan
    Button (655,128 62x28), "Stop"
        OnMouseClick: toggle Global.Tank1.Filling.Cmd.StopMan
    Button (720,128 62x28), "Resume"
        OnMouseClick: toggle Global.Tank1.Filling.Cmd.ResumeMan
    Rectangle (787,96 151x28), "Fill Lvl: %.2f m", text variable: Global.Tank1.Filling.ParamFillLevel
        OnMouseClick: write the text variable via Default
    Rectangle (787,128 89x28), "Act: %.2f m", text variable: Global.Tank1.Filling.WaterLevel
    Button (880,128 58x28), "Res.Done"
        OnMouseClick: toggle Global.Tank1.Filling.Cmd.ResetDone
    Rectangle (970,8 294x158)
    Label (974,10 140x18), "Phase: Draining"
    Button (975,32 50x26), "AUT"
        OnMouseClick: toggle Global.Tank1.Draining.Cmd.AutCtrl
    Button (1028,32 50x26), "MAN"
        OnMouseClick: toggle Global.Tank1.Draining.Cmd.ManCtrl
    Label (1086,36 38x18), "Idle"
    Label (1128,36 38x18), "Run"
    Label (1166,36 52x18), "Pause"
    Label (1218,36 44x18), "Done"
    Lamp1 (986,62 27x26), variable: Global.Tank1.Draining.State.AutCtrl, style: Lamp-Lamp1-Yellow
    Lamp1 (1039,62 27x26), variable: Global.Tank1.Draining.State.ManCtrl, style: Lamp-Lamp1-Yellow
    Lamp1 (1089,62 27x26), variable: Global.Tank1.Draining.State.Idle, style: Lamp-Lamp1-Yellow
    Lamp1 (1131,62 27x26), variable: Global.Tank1.Draining.State.Running, style: Lamp-Lamp1-Yellow
    Lamp1 (1177,62 27x26), variable: Global.Tank1.Draining.State.Paused, style: Lamp-Lamp1-Yellow
    Lamp1 (1224,62 27x26), variable: Global.Tank1.Draining.State.Done, style: Lamp-Lamp1-Yellow
    Button (975,96 62x28), "Start"
        OnMouseClick: toggle Global.Tank1.Draining.Cmd.StartMan
    Button (1040,96 62x28), "Pause"
        OnMouseClick: toggle Global.Tank1.Draining.Cmd.PauseMan
    Button (975,128 62x28), "Stop"
        OnMouseClick: toggle Global.Tank1.Draining.Cmd.StopMan
    Button (1040,128 62x28), "Resume"
        OnMouseClick: toggle Global.Tank1.Draining.Cmd.ResumeMan
    Rectangle (1107,96 151x28), "Drain Lvl: %.2f m", text variable: Global.Tank1.Draining.ParamDrainLevel
        OnMouseClick: write the text variable via Default
    Rectangle (1107,128 89x28), "Act: %.2f m", text variable: Global.Tank1.Draining.WaterLevel
    Button (1200,128 58x28), "Res.Done"
        OnMouseClick: toggle Global.Tank1.Draining.Cmd.ResetDone
    Rectangle (650,188 294x158)
    Label (654,190 140x18), "Phase: Mixing"
    Button (655,212 50x26), "AUT"
        OnMouseClick: toggle Global.Tank1.Mixing.Cmd.AutCtrl
    Button (708,212 50x26), "MAN"
        OnMouseClick: toggle Global.Tank1.Mixing.Cmd.ManCtrl
    Label (766,216 38x18), "Idle"
    Label (808,216 38x18), "Run"
    Label (846,216 52x18), "Pause"
    Label (898,216 44x18), "Done"
    Lamp1 (666,242 27x26), variable: Global.Tank1.Mixing.State.AutCtrl, style: Lamp-Lamp1-Yellow
    Lamp1 (719,242 27x26), variable: Global.Tank1.Mixing.State.ManCtrl, style: Lamp-Lamp1-Yellow
    Lamp1 (769,242 27x26), variable: Global.Tank1.Mixing.State.Idle, style: Lamp-Lamp1-Yellow
    Lamp1 (811,242 27x26), variable: Global.Tank1.Mixing.State.Running, style: Lamp-Lamp1-Yellow
    Lamp1 (857,242 27x26), variable: Global.Tank1.Mixing.State.Paused, style: Lamp-Lamp1-Yellow
    Lamp1 (904,242 27x26), variable: Global.Tank1.Mixing.State.Done, style: Lamp-Lamp1-Yellow
    Button (655,276 62x28), "Start"
        OnMouseClick: toggle Global.Tank1.Mixing.Cmd.StartMan
    Button (720,276 62x28), "Pause"
        OnMouseClick: toggle Global.Tank1.Mixing.Cmd.PauseMan
    Button (655,308 62x28), "Stop"
        OnMouseClick: toggle Global.Tank1.Mixing.Cmd.StopMan
    Button (720,308 62x28), "Resume"
        OnMouseClick: toggle Global.Tank1.Mixing.Cmd.ResumeMan
    Rectangle (787,276 151x28), "Mix Time: %d s", text variable: Global.Tank1.Mixing.ParamTimeSec
        OnMouseClick: write the text variable via Default
    Rectangle (787,308 89x28), "Elap: %d s", text variable: Global.Tank1.Mixing.ElapsedTimeSec
    Button (880,308 58x28), "Res.Done"
        OnMouseClick: toggle Global.Tank1.Mixing.Cmd.ResetDone
    Rectangle (970,188 294x158)
    Label (974,190 140x18), "Phase: Heating"
    Button (975,212 50x26), "AUT"
        OnMouseClick: toggle Global.Tank1.Heating.Cmd.AutCtrl
    Button (1028,212 50x26), "MAN"
        OnMouseClick: toggle Global.Tank1.Heating.Cmd.ManCtrl
    Label (1086,216 38x18), "Idle"
    Label (1128,216 38x18), "Run"
    Label (1166,216 52x18), "Pause"
    Label (1218,216 44x18), "Done"
    Lamp1 (986,242 27x26), variable: Global.Tank1.Heating.State.AutCtrl, style: Lamp-Lamp1-Yellow
    Lamp1 (1039,242 27x26), variable: Global.Tank1.Heating.State.ManCtrl, style: Lamp-Lamp1-Yellow
    Lamp1 (1089,242 27x26), variable: Global.Tank1.Heating.State.Idle, style: Lamp-Lamp1-Yellow
    Lamp1 (1131,242 27x26), variable: Global.Tank1.Heating.State.Running, style: Lamp-Lamp1-Yellow
    Lamp1 (1177,242 27x26), variable: Global.Tank1.Heating.State.Paused, style: Lamp-Lamp1-Yellow
    Lamp1 (1224,242 27x26), variable: Global.Tank1.Heating.State.Done, style: Lamp-Lamp1-Yellow
    Button (975,276 62x28), "Start"
        OnMouseClick: toggle Global.Tank1.Heating.Cmd.StartMan
    Button (1040,276 62x28), "Pause"
        OnMouseClick: toggle Global.Tank1.Heating.Cmd.PauseMan
    Button (975,308 62x28), "Stop"
        OnMouseClick: toggle Global.Tank1.Heating.Cmd.StopMan
    Button (1040,308 62x28), "Resume"
        OnMouseClick: toggle Global.Tank1.Heating.Cmd.ResumeMan
    Rectangle (1107,276 151x28), "Req Temp: %.1f C", text variable: Global.Tank1.Heating.ParamReqTemp
        OnMouseClick: write the text variable via Default
    Rectangle (1107,308 89x28), "Hold: %d s", text variable: Global.Tank1.Heating.fTime
    Button (1200,308 58x28), "Res.Done"
        OnMouseClick: toggle Global.Tank1.Heating.Cmd.ResetDone
    Rectangle (8,425 810x78)
    Label (16,429 180x20), "Batch Automat (Test)"
    Button (18,456 105x34), "Start Batch"
        OnMouseClick: toggle Test.bStartBatch
    Button (133,456 105x34), "Stop Batch"
        OnMouseClick: toggle Test.bStopBatch
    Label (255,436 38x18), "Run"
    Lamp1 (257,460 27x26), variable: Test.bRunning, style: Lamp-Lamp1-Yellow
    Rectangle (310,456 150x34), "Batches: %d", text variable: Test.nTargetBatches
        OnMouseClick: write the text variable via Default
    Rectangle (475,456 150x34), "Done: %d", text variable: Test.nCompletedBatches
    Rectangle (640,456 150x34), "Step: %d", text variable: Test.State
END_VISUALIZATION
